// TwinCAT 3 PLC project Biegbert_SPS
// ProgramVersion: 3.1.4026.27
// CompilerDefines: SIM
// libraries:
//   Tc2_MC2, * (Beckhoff Automation GmbH)
//   Tc2_MC2_Camming, * (Beckhoff Automation GmbH)
//   Tc2_Standard, * (Beckhoff Automation GmbH)
//   Tc2_System, * (Beckhoff Automation GmbH)
//   TcUnit, * (www.tcunit.org)
// project tree:
//   07_Test/ FB_BendKinematics_Test.TcPOU, PRG_TEST.TcPOU
//   00_GVL/ GVL_Config.TcGVL, GVL_HMI.TcGVL, GVL_Axis.TcGVL, GVL_Devices.TcGVL, GVL_IO.TcGVL, GVL_Plan.TcGVL, GVL_Sim.TcGVL
//   01_DUT/ E_AlarmCode.TcDUT, E_AlarmSeverity.TcDUT, E_Axis.TcDUT, E_AxisState.TcDUT, E_ClampState.TcDUT, E_CmdResult.TcDUT, E_HmiCmd.TcDUT, E_KinState.TcDUT, E_MotionMode.TcDUT, E_OperatingMode.TcDUT, ST_AlarmEntry.TcDUT, ST_HmiAlarms.TcDUT, ST_HmiAxisStatus.TcDUT, ST_HmiClampStatus.TcDUT, ST_HmiCmd.TcDUT, ST_HmiCmdAck.TcDUT, ST_HmiIoStatus.TcDUT, ST_HmiJog.TcDUT, ST_HmiParam.TcDUT, ST_HmiStatus.TcDUT, ST_KinStatus.TcDUT, ST_Material.TcDUT, E_G0Step.TcDUT, E_G2Step.TcDUT, E_G3Step.TcDUT, ST_FeedPoint.TcDUT, ST_PlanHeader.TcDUT, ST_PlanPoint.TcDUT, ST_PlanSection.TcDUT, ST_PlanTransfer.TcDUT, ST_RotPoint.TcDUT
//   04_Kinematics/ FB_BendKinematics.TcPOU, I_Kinematics.TcIO, F_ChuckInZone.TcPOU, F_ClampBlocking.TcPOU, F_Z1Max.TcPOU
//   02_IO/ FB_IoMap.TcPOU, FB_IoSim.TcPOU
//   03_Devices/ FB_Axis.TcPOU, FB_Clamp.TcPOU, F_Mod360.TcPOU
//   05_Sequence/ FB_BendSequence.TcPOU, FB_Interlocks.TcPOU, FB_ModeManager.TcPOU
//   06_HMI/ FB_AlarmManager.TcPOU, FB_HmiCommand.TcPOU, FB_HmiStatus.TcPOU, FB_PlanStore.TcPOU, F_PlanChecksum.TcPOU
//   / PlcTask.TcTTO
//   POUs/ MAIN.TcPOU
// real-time tasks:
//   TASK PlcTask: cycle T#10ms, priority 20, ADS port 350
// motion (NC):
//   TASK NC-Task 1 SAF: cycle T#2ms, priority 4, ADS port 501
//   TASK NC-Task 1 SVB: cycle T#10ms, priority 8, ADS port 511
//   AXIS Z1 (id 1)
//     Dynamic: AccelerationMaximum=200, DecelerationMaximum=200, Acceleration=200, Deceleration=200
//     Velo: Maximum=50
//     OtherSettings: AllowMotionCmdToSlave=true
//     encoder EncType=1
//       SoftEndMinControl: Enable=true, Range=-30
//       SoftEndMaxControl: Enable=true, Range=1282
//     drive DrvType=5
//       Analog: VeloReferenz=100, TorqueSetpointScale=10, ScaleFactorActTorque=0.1
//       TimeComp: TaskDelayCycles=1
//     controller CtrType=1
//       CtrPara: PriorControlFactor=1
//         Observer: BandWidth=20
//   AXIS Z2 (id 2)
//     Dynamic: AccelerationMaximum=100, DecelerationMaximum=100, Acceleration=100, Deceleration=100
//     Velo: Maximum=28.6
//     OtherSettings: AllowMotionCmdToSlave=true
//     encoder EncType=1
//       SoftEndMinControl: Enable=true, Range=-50
//       SoftEndMaxControl: Enable=true, Range=48
//     drive DrvType=5
//       Analog: VeloReferenz=57.2, TorqueSetpointScale=10, ScaleFactorActTorque=0.1
//     controller CtrType=1
//       CtrPara: PriorControlFactor=1
//         Observer: BandWidth=20
//   AXIS X (id 3)
//     Dynamic: AccelerationMaximum=20, DecelerationMaximum=20, Acceleration=20, Deceleration=20
//     Velo: Maximum=3.5
//     OtherSettings: AllowMotionCmdToSlave=true
//     encoder EncType=1
//       SoftEndMinControl: Enable=true, Range=-50
//       SoftEndMaxControl: Enable=true, Range=50
//     drive DrvType=5
//       Analog: VeloReferenz=7, TorqueSetpointScale=10, ScaleFactorActTorque=0.1
//     controller CtrType=1
//       CtrPara: PriorControlFactor=1
//         Observer: BandWidth=20
//   AXIS A (id 4)
//     General: UnitName=°
//     Dynamic: AccelerationMaximum=360, DecelerationMaximum=360, Acceleration=360, Deceleration=360
//     Velo: Maximum=180
//     OtherSettings: AllowMotionCmdToSlave=true
//     encoder EncType=1
//       SoftEndMinControl: Enable=true, Range=-60
//       SoftEndMaxControl: Enable=true, Range=60
//     drive DrvType=5
//       Analog: VeloReferenz=360, TorqueSetpointScale=10, ScaleFactorActTorque=0.1
//     controller CtrType=1
//       CtrPara: PriorControlFactor=1
//         Observer: BandWidth=20
//   AXIS W (id 5)
//     Dynamic: AccelerationMaximum=360, DecelerationMaximum=360, Acceleration=360, Deceleration=360
//     Velo: Maximum=180
//     OtherSettings: AllowMotionCmdToSlave=true
//     encoder EncType=1
//     drive DrvType=5
//       Analog: VeloReferenz=360, TorqueSetpointScale=10, ScaleFactorActTorque=0.1
//     controller CtrType=1
//       CtrPara: PriorControlFactor=1
//         Observer: BandWidth=20
// variable links:
//   (this object) <-> NC-Task 1 SAF/Axes/A
//     PlcTask Inputs/GVL_Axis.A.NcToPlc <-> Outputs/ToPlc
//     PlcTask Outputs/GVL_Axis.A.PlcToNc <-> Inputs/FromPlc
//   (this object) <-> NC-Task 1 SAF/Axes/W
//     PlcTask Inputs/GVL_Axis.W.NcToPlc <-> Outputs/ToPlc
//     PlcTask Outputs/GVL_Axis.W.PlcToNc <-> Inputs/FromPlc
//   (this object) <-> NC-Task 1 SAF/Axes/X
//     PlcTask Inputs/GVL_Axis.X.NcToPlc <-> Outputs/ToPlc
//     PlcTask Outputs/GVL_Axis.X.PlcToNc <-> Inputs/FromPlc
//   (this object) <-> NC-Task 1 SAF/Axes/Z1
//     PlcTask Inputs/GVL_Axis.Z1.NcToPlc <-> Outputs/ToPlc
//     PlcTask Outputs/GVL_Axis.Z1.PlcToNc <-> Inputs/FromPlc
//   (this object) <-> NC-Task 1 SAF/Axes/Z2
//     PlcTask Inputs/GVL_Axis.Z2.NcToPlc <-> Outputs/ToPlc
//     PlcTask Outputs/GVL_Axis.Z2.PlcToNc <-> Inputs/FromPlc

CONFIGURATION Biegbert_SPS
    RESOURCE PLC ON TwinCAT3
        TASK PlcTask(INTERVAL := T#10ms, PRIORITY := 20);
        PROGRAM MAIN WITH PlcTask : MAIN;
    END_RESOURCE
END_CONFIGURATION

// ---- 01_DUT/E_AlarmCode.TcDUT
// Alarmcodes. Die Texte liegen im Backend (backend/biegbert/alarms.py).
{attribute 'qualified_only'}
{attribute 'strict'}
{attribute 'to_string'}
TYPE E_AlarmCode :
(
    None := 0,
    HmiHeartbeatLost := 1001, // Heartbeat ausgefallen
    SimulationActive := 1002, // Simulationsbetrieb aktiv
    EStopActive := 1100, // Not-Halt ausgelöst
    SafetyNotReady := 1101, // TwinSAFE nicht betriebsbereit
    AxisError := 2000, // nSource = E_Axis, nDetail = NC-Fehlercode
    AxisLagError := 2001, // Schleppfehler
    AxisSoftLimit := 2002, // Software-Endlage
    AxisTorqueLimit := 2003, // Momentgrenze
    ClampTimeout := 3000, // nSource = Niederhalter
    ClampPressureLow := 3001, // Klemmdruck fehlt
    ClampZoneViolation := 3002, // 4BF-Zone bei geschlossenem Niederhalter
    DistanceZ1Z2 := 4000, // dZ12 unterschritten
    KinCoupleFailed := 5000, // Kopplung oder Kurvenscheibe fehlgeschlagen, nDetail = NC-Fehlercode
    KinMasterFault := 5001, // Master Z1 gestört
    KinSlaveFault := 5002, // Slave gestört
    KinPositionDeviation := 5003, // Achse weicht vor Wiederanlauf vom Plan ab
    SeqStepTimeout := 6001 // Schritt hängt, nDetail = Schrittnummer
) UDINT;
END_TYPE

// ---- 01_DUT/E_AlarmSeverity.TcDUT
// Abgestufte Reaktion nach SE3.
{attribute 'qualified_only'}
{attribute 'strict'}
{attribute 'to_string'}
TYPE E_AlarmSeverity :
(
    None := 0,
    Info := 1, // nur Anzeige
    Warning := 2, // Anzeige, Ablauf läuft weiter
    Stop := 3, // Pause
    Fault := 4 // Pause, Wiederanlauf erst nach Behebung
) INT;
END_TYPE

// ---- 01_DUT/E_Axis.TcDUT
// Achsen. Die Werte sind die Indizes von aAxis in ST_HmiStatus.
{attribute 'qualified_only'}
{attribute 'strict'}
{attribute 'to_string'}
TYPE E_Axis :
(
    None := 0, // keine Achse
    Z1 := 1, // Vorschub, mm
    Z2 := 2, // Führung, mm
    X := 3, // Matrizenauslenkung, mm
    A := 4, // Matrizendrehung, °
    W := 5 // Rohrdrehung, °, Modulo
) INT;
END_TYPE

// ---- 01_DUT/E_AxisState.TcDUT
// Vereinfachter Achszustand für die GUI.
{attribute 'qualified_only'}
{attribute 'strict'}
{attribute 'to_string'}
TYPE E_AxisState :
(
    Disabled := 0,
    Standstill := 1,
    Moving := 2, // Einzelbewegung
    Coupled := 3, // über FB_BendKinematics gekoppelt
    Error := 4
) INT;
END_TYPE

// ---- 01_DUT/E_ClampState.TcDUT
// Zustand eines Niederhalters.
{attribute 'qualified_only'}
{attribute 'strict'}
{attribute 'to_string'}
TYPE E_ClampState :
(
    Unknown := 0,
    Open := 1, // Endlage OFFEN gemeldet
    Closing := 2, // Ventil an, Schaltzeit läuft
    Clamped := 3, // OFFEN verlassen, Druck ok, Schaltzeit abgelaufen
    Opening := 4, // Ventil aus, Endlage noch nicht erreicht
    Fault := 5 // Zeitüberwachung oder Plausibilität verletzt
) INT;
END_TYPE

// ---- 01_DUT/E_CmdResult.TcDUT
// Ergebnis der Kommandoprüfung.
{attribute 'qualified_only'}
{attribute 'strict'}
{attribute 'to_string'}
TYPE E_CmdResult :
(
    None := 0, // noch keine Antwort
    Accepted := 1, // angenommen, Ausführung siehe Status
    RejectedUnknown := 2, // Kommando unbekannt
    RejectedMode := 3, // in dieser Betriebsart nicht erlaubt
    RejectedInterlock := 4, // Verriegelung aktiv
    RejectedParam := 5, // Parameter ungültig
    RejectedSequence := 6, // zweite Stufe ohne gültige erste Stufe
    RejectedBusy := 7 // Gerät beschäftigt
) INT;
END_TYPE

// ---- 01_DUT/E_HmiCmd.TcDUT
// Kommandos der GUI. Details: docs/hmi-schnittstelle.md
{attribute 'qualified_only'}
{attribute 'strict'}
{attribute 'to_string'}
TYPE E_HmiCmd :
(
    None := 0,
    AlarmAck := 10, // nValue = Alarm-Slot, 0 = alle
    ParamApply := 11, // stParam prüfen und übernehmen
    AxisEnable := 100, // Phase 4/6: eAxis
    AxisDisable := 101, // Phase 6: eAxis
    AxisReset := 102, // Phase 6: eAxis
    AxisHalt := 103, // Phase 4/6: eAxis
    AxisMoveAbs := 104, // Phase 6: eAxis, fPosition, fVelocity
    ClampOpen := 120, // Phase 6: nClamp
    ClampClose := 121, // Phase 6: nClamp
    ModePause := 200, // Phase 6
    ModeResume1 := 201, // Phase 6: RES1
    ModeResume2 := 202, // Phase 6: RES2
    ModeSingleAxis1 := 203, // Phase 6: MAN1
    ModeSingleAxis2 := 204, // Phase 6: MAN2
    ModeReturnToBase := 205, // Phase 6: OK, nur bei GZ_POS
    SimSetInput := 300, // Phase 5/6: nur im Simulationsbetrieb, nValue = Signal-ID, fPosition <> 0 = TRUE
    SimInjectFault := 301, // Phase 5: nur im Simulationsbetrieb, nValue = Fehler-ID
    SeqStart := 400, // reserviert Phase 8: ST
    SeqConfirmQ1 := 401, // reserviert Phase 8
    SeqConfirmQ2 := 402, // reserviert Phase 8
    SeqPartRemoved := 403, // reserviert Phase 8: ENT
    PlanLoad := 410, // reserviert Phase 9
    MaterialConfirm := 411, // reserviert Phase 9
    CalibrateAxis := 500 // reserviert Phase 9: Einmessen
) UDINT;
END_TYPE

// ---- 01_DUT/E_KinState.TcDUT
// Zustand der Kinematik.
{attribute 'qualified_only'}
{attribute 'strict'}
{attribute 'to_string'}
TYPE E_KinState :
(
    Idle := 0, // kein Plan aktiv
    Loaded := 1, // Plan geladen, entkoppelt
    Coupling := 2,
    Running := 3, // gekoppelt, Master läuft
    Holding := 4, // Master bremst
    Held := 5, // gekoppelt, Stillstand
    Decoupling := 6,
    Fault := 7 // Reset nötig
) INT;
END_TYPE

// ---- 01_DUT/E_MotionMode.TcDUT
// Bewegungsmodus der Kinematik.
{attribute 'qualified_only'}
{attribute 'strict'}
{attribute 'to_string'}
TYPE E_MotionMode :
(
    Single := 1, // entkoppelt, Einzelachsen erlaubt
    Coupled := 2, // gekoppelt, Master läuft oder fährt an
    Hold := 3 // gekoppelt, Master hält
) INT;
END_TYPE

// ---- 01_DUT/E_OperatingMode.TcDUT
// Betriebsart. Die Werte entsprechen den GRAFCET-Schritten von G1.
{attribute 'qualified_only'}
{attribute 'strict'}
{attribute 'to_string'}
TYPE E_OperatingMode :
(
    Automatic := 10, // G1 Schritt 10
    Pause := 11, // G1 Schritt 11
    SingleAxis := 12, // G1 Schritt 12
    ReturnToBase := 13 // G1 Schritt 13
) INT;
END_TYPE

// ---- 01_DUT/ST_AlarmEntry.TcDUT
// Ein Alarm. Texte und Historie liegen im Backend.
{attribute 'pack_mode' := '1'}
TYPE ST_AlarmEntry :
STRUCT
    eCode : E_AlarmCode;
    eSeverity : E_AlarmSeverity;
    nSource : DINT; // Achse oder Niederhalter
    nDetail : UDINT;
    nTimestamp : ULINT; // Windows-Dateizeit, 100 ns
    bActive : BOOL; // Ursache besteht noch
    bAcked : BOOL;
END_STRUCT
END_TYPE

// ---- 01_DUT/ST_HmiAlarms.TcDUT
// SPS -> GUI. Aktive oder nicht quittierte Alarme.
{attribute 'pack_mode' := '1'}
TYPE ST_HmiAlarms :
STRUCT
    nChangeCounter : UDINT; // bei jeder Änderung +1
    nCount : UINT;
    bOverflow : BOOL;
    eHighestSeverity : E_AlarmSeverity;
    aEntry : ARRAY[1..32] OF ST_AlarmEntry;
END_STRUCT
END_TYPE

// ---- 01_DUT/ST_HmiAxisStatus.TcDUT
// SPS -> GUI. Status einer Achse.
{attribute 'pack_mode' := '1'}
TYPE ST_HmiAxisStatus :
STRUCT
    eState : E_AxisState;
    bEnabled : BOOL;
    bReady : BOOL;
    bError : BOOL;
    nErrorId : UDINT;
    fActPos : LREAL; // mm oder °
    fSetPos : LREAL;
    fActVelo : LREAL; // mm/s oder °/s
    fSetVelo : LREAL;
    fLagError : LREAL; // mm oder °
    fTorque_Nm : LREAL;
END_STRUCT
END_TYPE

// ---- 01_DUT/ST_HmiClampStatus.TcDUT
// SPS -> GUI. Status eines Niederhalters.
{attribute 'pack_mode' := '1'}
TYPE ST_HmiClampStatus :
STRUCT
    eState : E_ClampState;
    bValve : BOOL; // Ausgang
    bOpen : BOOL; // Endlage OFFEN
    fLastSwitchTime_ms : LREAL;
END_STRUCT
END_TYPE

// ---- 01_DUT/ST_HmiCmd.TcDUT
// GUI -> SPS. Die GUI schreibt hier, die SPS liest nur.
{attribute 'pack_mode' := '1'}
TYPE ST_HmiCmd :
STRUCT
    nHeartbeat : UDINT; // alle 100 ms hochzählen
    nCmdId : UDINT; // zuletzt und getrennt schreiben
    eCmd : E_HmiCmd;
    eAxis : E_Axis;
    nClamp : USINT; // 1..6, 0 = keiner
    fPosition : LREAL; // mm oder °, je nach Achse
    fVelocity : LREAL; // mm/s oder °/s
    nValue : DINT; // kommandoabhängig
    stJog : ST_HmiJog;
END_STRUCT
END_TYPE

// ---- 01_DUT/ST_HmiCmdAck.TcDUT
// SPS -> GUI. Antwort auf das letzte Kommando.
{attribute 'pack_mode' := '1'}
TYPE ST_HmiCmdAck :
STRUCT
    nAckId : UDINT; // gleich nCmdId, sobald geprüft
    eResult : E_CmdResult;
    nDetail : UDINT; // z. B. fehlende Bedingung
END_STRUCT
END_TYPE

// ---- 01_DUT/ST_HmiIoStatus.TcDUT
// SPS -> GUI. E/A-Übersicht ohne Niederhalter. Belegung folgt mit der EMSR-Liste.
{attribute 'pack_mode' := '1'}
TYPE ST_HmiIoStatus :
STRUCT
    bPressureOk : BOOL; // Druckschalter SDE5
    abPanelIn : ARRAY[1..16] OF BOOL; // ED1809
    abPanelOut : ARRAY[1..16] OF BOOL; // ED2809
END_STRUCT
END_TYPE

// ---- 01_DUT/ST_HmiJog.TcDUT
// Tippen. Wird zyklisch ausgewertet und läuft nicht über den Handshake.
{attribute 'pack_mode' := '1'}
TYPE ST_HmiJog :
STRUCT
    eAxis : E_Axis;
    nDirection : SINT; // -1, 0, +1
    fVelocityFactor_pct : LREAL; // 0..100 der Einrichtgeschwindigkeit
END_STRUCT
END_TYPE

// ---- 01_DUT/ST_HmiParam.TcDUT
// GUI -> SPS mit Übernahme durch ParamApply.
{attribute 'pack_mode' := '1'}
TYPE ST_HmiParam :
STRUCT
    nPlanId : UDINT;
    stMaterial : ST_Material;
    fFeedOverride_pct : LREAL; // 0..100
    fSingleAxisVelo_pct : LREAL; // 0..100
END_STRUCT
END_TYPE

// ---- 01_DUT/ST_HmiStatus.TcDUT
// SPS -> GUI. Die SPS schreibt hier, die GUI liest nur.
{attribute 'pack_mode' := '1'}
TYPE ST_HmiStatus :
STRUCT
    nLifeCounter : UDINT; // pro SPS-Zyklus +1
    bHmiAlive : BOOL;
    bSimulation : BOOL;
    bEStopActive : BOOL;
    bSafetyOk : BOOL;
    eMode : E_OperatingMode;
    nStepG2 : INT; // GRAFCET-Schritt
    nStepG3 : INT;
    nBend : UDINT; // aktueller Bogen
    dwBaseStateMissing : DWORD; // Bitmaske, siehe Doku
    stCmdAck : ST_HmiCmdAck;
    aAxis : ARRAY[1..5] OF ST_HmiAxisStatus; // Index = E_Axis
    aClamp : ARRAY[1..6] OF ST_HmiClampStatus;
    stIo : ST_HmiIoStatus;
    stKin : ST_KinStatus;
    stParamActive : ST_HmiParam;
END_STRUCT
END_TYPE

// ---- 01_DUT/ST_KinStatus.TcDUT
// Status von I_Kinematics.
{attribute 'pack_mode' := '1'}
TYPE ST_KinStatus :
STRUCT
    eState : E_KinState;
    eMode : E_MotionMode;
    nPlanId : UDINT;
    bError : BOOL;
    nErrorId : UDINT;
    fMasterPos_mm : LREAL;
END_STRUCT
END_TYPE

// ---- 01_DUT/ST_Material.TcDUT
// Halbzeugdaten des aktiven Programms.
{attribute 'pack_mode' := '1'}
TYPE ST_Material :
STRUCT
    fDiameter_mm : LREAL;
    fWall_mm : LREAL; // 0 = Vollmaterial
    fYield_MPa : LREAL; // Rp0,2
    fForceLimit_N : LREAL;
END_STRUCT
END_TYPE

// ---- 01_DUT/E_G0Step.TcDUT
// GRAFCET G0 Not-Halt [Langfeld].
{attribute 'qualified_only'}
{attribute 'strict'}
{attribute 'to_string'}
TYPE E_G0Step :
(
    S1_Betrieb := 1,
    S2_NotHalt := 2
) INT;
END_TYPE

// ---- 01_DUT/E_G2Step.TcDUT
// GRAFCET G2 Biegevorgang [Langfeld], Nummern = GRAFCET-Schritte.
{attribute 'qualified_only'}
{attribute 'strict'}
{attribute 'to_string'}
TYPE E_G2Step :
(
    S20_Grundzustand := 20,      // wartet auf Start
    S21_Startposition := 21,     // Z2, X, A und Z1 auf Startposition des Abschnitts
    S22_Niederhalter := 22,      // NH_soll schließen, Klemmung prüfen
    S23_Biegen := 23,            // gekoppelt: Z1 Master, X und A aus Kurvenscheibe
    S24_Halten := 24,            // Geometrie unter Last halten, warten auf Q1
    S25_NhOeffnen := 25,         // alle Niederhalter öffnen, warten auf Q2
    S26_Neutral := 26,           // entkoppeln, X und A auf 0
    S27_Uebergabe := 27,         // n := n + 1; weiterer Abschnitt oder warten auf ENT / Fortsetzung
    S28_Grundstellung := 28      // Z1, Z2, W auf 0
) INT;
END_TYPE

// ---- 01_DUT/E_G3Step.TcDUT
// GRAFCET G3 Werkstückrotation [Langfeld].
{attribute 'qualified_only'}
{attribute 'strict'}
{attribute 'to_string'}
TYPE E_G3Step :
(
    S30_Bereit := 30,
    S31_Stop := 31,     // Master steht an der Rotationsposition
    S32_Drehen := 32    // W dreht
) INT;
END_TYPE

// ---- 01_DUT/ST_FeedPoint.TcDUT
// Ab Z1-Position fZ1_mm gilt der Vorschub fFeed_mm_s.
{attribute 'pack_mode' := '1'}
TYPE ST_FeedPoint :
STRUCT
    fZ1_mm : LREAL;
    fFeed_mm_s : LREAL;
END_STRUCT
END_TYPE

// ---- 01_DUT/ST_PlanHeader.TcDUT
{attribute 'pack_mode' := '1'}
TYPE ST_PlanHeader :
STRUCT
    nPlanId : UDINT;
    nFormat : UINT;           // = GVL_Config.cPlanFormat
    nSectionCount : UINT;
    nPointCount : UDINT;
    nChecksum : UDINT;        // F_PlanChecksum über die belegten Abschnitte und Punkte
    stMaterial : ST_Material;
END_STRUCT
END_TYPE

// ---- 01_DUT/ST_PlanPoint.TcDUT
// Stützpunkt der Kurvenscheibe: Masterposition s (= Z1) mit u (= X) und phi (= A).
{attribute 'pack_mode' := '1'}
TYPE ST_PlanPoint :
STRUCT
    fS_mm : LREAL;
    fU_mm : LREAL;
    fPhi_deg : LREAL;
END_STRUCT
END_TYPE

// ---- 01_DUT/ST_PlanSection.TcDUT
// Ein Abschnitt = eine Kurvenscheibe mit konstantem Z2. Geraden sind Teil der Kurvenscheibe (u = 0).
{attribute 'pack_mode' := '1'}
TYPE ST_PlanSection :
STRUCT
    fZ1Start_mm : LREAL;
    fZ1Fin_mm : LREAL;
    fZ2_mm : LREAL;
    nFirstPoint : UDINT;      // Index in aPoint (1-basiert)
    nPointCount : UDINT;
    nFeedCount : UINT;
    aFeed : ARRAY[1..8] OF ST_FeedPoint;     // = GVL_Config.cMaxFeed
    nRotCount : UINT;
    aRot : ARRAY[1..16] OF ST_RotPoint;      // = GVL_Config.cMaxRot
    nClampMask : BYTE;        // Bit 0..5: NH1..NH6 zu Beginn schließen
    aClampOpen_mm : ARRAY[1..6] OF LREAL;    // Z1-Position, ab der NH i geöffnet wird
END_STRUCT
END_TYPE

// ---- 01_DUT/ST_PlanTransfer.TcDUT
// Übergabebereich Biegeplan (GVL_HMI.stPlanXfer) und aktiver Plan (GVL_Plan.stActive). 103552 Byte.
{attribute 'pack_mode' := '1'}
TYPE ST_PlanTransfer :
STRUCT
    stHeader : ST_PlanHeader;
    aSection : ARRAY[1..16] OF ST_PlanSection;    // = GVL_Config.cMaxSections
    aPoint : ARRAY[1..4000] OF ST_PlanPoint;      // = GVL_Config.cMaxPoints
END_STRUCT
END_TYPE

// ---- 01_DUT/ST_RotPoint.TcDUT
// Rotation von W um fW_deg (relativ), wenn Z1 fZ1_mm erreicht.
{attribute 'pack_mode' := '1'}
TYPE ST_RotPoint :
STRUCT
    fZ1_mm : LREAL;
    fW_deg : LREAL;
END_STRUCT
END_TYPE

// ---- 00_GVL/GVL_Config.TcGVL
// Feste Konfigurationswerte. Werte mit VORLÄUFIG stammen aus Doku/CAD und werden an der Anlage ersetzt.
// Gleiche Werte stehen im Backend in backend/biegbert/config.py (siehe 04_Datenfluss_und_Zustaende, Kap. 6).
{attribute 'qualified_only'}
VAR_GLOBAL CONSTANT
    cAxisCount           : INT  := 5;
    cClampCount          : INT  := 6;
    cAlarmSlots          : INT  := 32;
    tHeartbeatTimeout    : TIME := T#500MS;
    tTwoStepConfirmation : TIME := T#10S;

    // Achsen, Index = E_Axis (1 Z1, 2 Z2, 3 X, 4 A, 5 W). VORLÄUFIG.
    // W ist in der NC eine Rundachse OHNE Modulo; die SPS rechnet die Anzeige auf 0..360°.
    aAxisMin        : ARRAY[1..5] OF LREAL := [-30.0, -50.0, -50.0, -60.0, -1.0E9];
    aAxisMax        : ARRAY[1..5] OF LREAL := [1282.0, 48.0, 50.0, 60.0, 1.0E9];
    aAxisVMax       : ARRAY[1..5] OF LREAL := [50.0, 28.6, 3.5, 180.0, 180.0];   // mm/s bzw. °/s
    aAxisVSetup     : ARRAY[1..5] OF LREAL := [30.0, 10.0, 3.5, 20.0, 30.0];    // Einrichtgeschwindigkeit bei 100 %
    aAxisAccel      : ARRAY[1..5] OF LREAL := [200.0, 100.0, 20.0, 360.0, 360.0];
    aRatedTorque_Nm : ARRAY[1..5] OF LREAL := [15.2, 1.2, 1.37, 2.38, 1.37];  // Motor-Nennmoment (Bezug von 0x6077), VORLÄUFIG
    fPosTol         : LREAL := 0.05;   // mm bzw. °

    // Prozessgeometrie (CAD-Auswertung 24.11.2026). VORLÄUFIG.
    fVAtZ2Zero_mm       : LREAL := 24.0;     // Werkzeugabstand v bei Z2 = 0
    fZ1CollisionBase_mm : LREAL := 743.25;   // Z1-Grenze Futter <-> Führung bei Z2 = 0
    // Z1-Bereich, in dem das Futter die Zone des Niederhalterpaares 1..3 berührt (Paar k = NH 2k-1, 2k)
    aClampZoneLo_mm : ARRAY[1..3] OF LREAL := [508.25, 278.5, 50.5];
    aClampZoneHi_mm : ARRAY[1..3] OF LREAL := [710.75, 481.0, 253.0];
    tClampSwitchSim : TIME := T#120MS;   // Schaltzeit im Simulationsmodell
    tClampSwitch    : TIME := T#120MS;   // Mindestzeit bis „geklemmt“ (DFM-50, an der Anlage messen)
    tClampTimeout   : TIME := T#1S;      // Zeitüberwachung Öffnen/Schließen

    fForceLimitMax_N : LREAL := 25000.0;

    // Planübergabe (muss zu backend/biegbert/plc/layout.py passen)
    cPlanFormat  : UINT := 1;
    cMaxSections : INT := 16;
    cMaxFeed     : INT := 8;
    cMaxRot      : INT := 16;
    cMaxPoints   : INT := 4000;
END_VAR

// ---- 00_GVL/GVL_HMI.TcGVL
// Einzige Schnittstelle zur GUI. Details: docs/hmi-schnittstelle.md
// Backend schreibt stCmd, stParam, stPlanXfer; die SPS schreibt stStatus und stAlarm.
{attribute 'qualified_only'}
VAR_GLOBAL
    stCmd      : ST_HmiCmd;
    stStatus   : ST_HmiStatus;
    stParam    : ST_HmiParam;
    stAlarm    : ST_HmiAlarms;
    stPlanXfer : ST_PlanTransfer;   // Übergabebereich Biegeplan, wird nur bei PlanLoad gelesen
END_VAR

// ---- 00_GVL/GVL_Axis.TcGVL
// NC-Achsen. Im System Manager unter MOTION > NC-Task > Achsen > (Achse) > Einstellungen > „Mit SPS verknüpfen“
// die passende Variable wählen: Z1 -> GVL_Axis.Z1 usw.
{attribute 'qualified_only'}
VAR_GLOBAL
    Z1 : AXIS_REF;   // Vorschub
    Z2 : AXIS_REF;   // Führung („Eisenschwein“)
    X  : AXIS_REF;   // Matrizenauslenkung
    A  : AXIS_REF;   // Matrizendrehung
    W  : AXIS_REF;   // Rohrdrehung
END_VAR

// ---- 00_GVL/GVL_Devices.TcGVL
// Geräteinstanzen. MAIN ruft sie zyklisch auf; Ablauf und HMI-Bausteine rufen nur ihre Methoden.
{attribute 'qualified_only'}
VAR_GLOBAL
    aAxis   : ARRAY[1..5] OF FB_Axis;    // Index = E_Axis
    aClamp  : ARRAY[1..6] OF FB_Clamp;
    fbKin   : FB_BendKinematics;
    fbAlarm : FB_AlarmManager;
END_VAR

// ---- 00_GVL/GVL_IO.TcGVL
// Prozessabbild und logische Signale. Nur 02_IO greift auf die AT-Variablen zu (architektur.md, Regel 5).
// Die AT-Variablen im System Manager mit den Klemmen verknüpfen (docs/twincat-einrichtung.md).
{attribute 'qualified_only'}
VAR_GLOBAL
    // ── Eingänge ──
    abClampOpenIn    AT %I* : ARRAY[1..6] OF BOOL;   // EP1008 Kanal 1..6: SMT-8M Endlage OFFEN, NH1..NH6
    bPressureOkIn    AT %I* : BOOL;                  // EP1008 Kanal 7: SDE5 Klemmdruck in Ordnung
    bSafetyOkIn      AT %I* : BOOL;                  // TwinSAFE -> Standard-SPS: Sicherheitskreis geschlossen, STO aufgehoben
    bEStopReleasedIn AT %I* : BOOL;                  // TwinSAFE -> Standard-SPS: Not-Halt entriegelt
    abPanelIn        AT %I* : ARRAY[1..16] OF BOOL;  // ED1809, Belegung offen
    anTorqueIn       AT %I* : ARRAY[1..5] OF INT;    // AX8000 Torque actual value (0x6077, 0,1 % Nennmoment), Index = E_Axis
    // ── Ausgänge ──
    abClampValveOut  AT %Q* : ARRAY[1..6] OF BOOL;   // EP2008 Kanal 1..6: Ventil NH1..NH6, TRUE = schließen
    abPanelOut       AT %Q* : ARRAY[1..16] OF BOOL;  // ED2809, Belegung offen
    bCameraTriggerOut AT %Q* : BOOL;                 // EL2252 Kanal 1 (später)

    // ── logische Signale (FB_IoMap) ──
    abClampOpen  : ARRAY[1..6] OF BOOL;
    bPressureOk  : BOOL;
    bSafetyOk    : BOOL;
    bEStopActive : BOOL;
    abPanel      : ARRAY[1..16] OF BOOL;
    afTorque_Nm  : ARRAY[1..5] OF LREAL;
    abClampValve : ARRAY[1..6] OF BOOL;
    abPanelLamp  : ARRAY[1..16] OF BOOL;
    bCameraTrigger : BOOL;
END_VAR

// ---- 00_GVL/GVL_Plan.TcGVL
// Geprüfte Kopie des aktiven Biegeplans. Schreibt nur FB_PlanStore, liest FB_BendKinematics und FB_BendSequence.
{attribute 'qualified_only'}
VAR_GLOBAL
    stActive : ST_PlanTransfer;
    bValid   : BOOL;
END_VAR

// ---- 00_GVL/GVL_Sim.TcGVL
// Eingriffe der Simulation. Wirkt nur, wenn das Projekt mit dem Compiler-Define SIM übersetzt wurde.
// Gesetzt über die Kommandos SimSetInput und SimInjectFault.
{attribute 'qualified_only'}
VAR_GLOBAL
    bPressureOk  : BOOL := TRUE;
    bEStop       : BOOL;
    abAxisFault  : ARRAY[1..5] OF BOOL;   // simulierter Achsfehler, Index = E_Axis
    abClampStuck : ARRAY[1..6] OF BOOL;   // Endlage OFFEN bleibt hängen
END_VAR

// ---- 04_Kinematics/I_Kinematics.TcIO
// Einzige Schnittstelle des Ablaufs zur Achskopplung. Details: docs/kinematik.md
INTERFACE I_Kinematics

METHOD Cyclic
// Einmal pro SPS-Zyklus aufrufen.
VAR_INPUT
END_VAR
END_METHOD

METHOD LoadPlan : BOOL
// Aktiven Plan (GVL_Plan.stActive) mit dieser ID übernehmen. Nur entkoppelt.
VAR_INPUT
    nPlanId : UDINT;
END_VAR
END_METHOD

METHOD LoadSection : BOOL
// Kurvenscheiben des Abschnitts nSection laden. Nur entkoppelt; fertig, wenn TableReady() TRUE meldet.
VAR_INPUT
    nSection : INT;
END_VAR
END_METHOD

METHOD TableReady : BOOL
VAR_INPUT
END_VAR
END_METHOD

METHOD Start : BOOL
// Koppelt X und A an Z1 und startet den Master.
VAR_INPUT
END_VAR
END_METHOD

METHOD Hold : BOOL
// Bremst den Master. Die Kopplung bleibt bestehen.
VAR_INPUT
END_VAR
END_METHOD

METHOD Resume : BOOL
// Setzt den Master aus dem Halt fort (nicht an einer offenen Rotation oder am Abschnittsende).
VAR_INPUT
END_VAR
END_METHOD

METHOD AtRotation : BOOL
// Master steht an einer Rotationsposition; RotationAngle() liefert den Drehwinkel für W.
VAR_INPUT
END_VAR
END_METHOD

METHOD RotationAngle : LREAL
VAR_INPUT
END_VAR
END_METHOD

METHOD ContinueAfterRotation : BOOL
VAR_INPUT
END_VAR
END_METHOD

METHOD SectionDone : BOOL
// Master steht am Ende des Abschnitts, Kopplung besteht noch.
VAR_INPUT
END_VAR
END_METHOD

METHOD Abort : BOOL
// Stoppt den Master und löst die Kopplung.
VAR_INPUT
END_VAR
END_METHOD

METHOD Reset : BOOL
// Quittiert einen Fehler der Kinematik. Der Plan bleibt erhalten.
VAR_INPUT
END_VAR
END_METHOD

METHOD Unload : BOOL
// Plan verwerfen (nur entkoppelt).
VAR_INPUT
END_VAR
END_METHOD

METHOD IsCoupled : BOOL
VAR_INPUT
END_VAR
END_METHOD

METHOD GetStatus : ST_KinStatus
VAR_INPUT
END_VAR
END_METHOD

END_INTERFACE

// ---- POUs/MAIN.TcPOU
PROGRAM MAIN
// Zyklusreihenfolge nach docs/architektur.md:
// 1 Eingänge, 2 Kommandos, 3 Abläufe, 4 Kinematik und Geräte, 5 Ausgänge, 6 Status und Alarme.
VAR
    fbIo : FB_IoMap;
    fbCmd : FB_HmiCommand;
    fbMode : FB_ModeManager;
    fbSeq : FB_BendSequence;
    fbPlan : FB_PlanStore;
    fbInterlocks : FB_Interlocks;
    fbStatus : FB_HmiStatus;
    dwBaseMissing : DWORD;
    bKinLock : BOOL;
    abSimFault : ARRAY[1..5] OF BOOL;
    bSim : BOOL;
    bInit : BOOL := TRUE;
    i : INT;
END_VAR

// 1 Eingänge
fbIo.ReadInputs();
bSim := fbIo.IsSimulation();
IF bInit THEN
    bInit := FALSE;
    IF bSim THEN
        GVL_Devices.fbAlarm.Raise(E_AlarmCode.SimulationActive, E_AlarmSeverity.Info, 0, 0);
    END_IF
END_IF
{IF defined (SIM)}
abSimFault := GVL_Sim.abAxisFault;
{END_IF}

// 2 Kommandos
dwBaseMissing := fbStatus.CalcBaseMissing(fbSeq.bMaterialOk);
fbCmd(fbMode := fbMode, fbSeq := fbSeq, fbPlan := fbPlan, dwBaseMissing := dwBaseMissing, bSimulation := bSim);

// 3 Abläufe
fbMode(bEStopActive := GVL_IO.bEStopActive, bSafetyOk := GVL_IO.bSafetyOk,
       nStopCounter := GVL_Devices.fbAlarm.nStopCounter);
fbSeq(bFree := fbMode.bFree, bAbort := fbMode.bEnteredSingle, bInit := fbMode.bInitSequences);

// 4 Kinematik und Geräte
GVL_Devices.fbKin.Cyclic();
bKinLock := GVL_Devices.fbKin.IsCoupled();
GVL_Devices.aAxis[1](pAxis := ADR(GVL_Axis.Z1), nIndex := 1, bAllowPower := NOT GVL_IO.bEStopActive,
    bLockedByKin := bKinLock, bSimFault := abSimFault[1], fTorque_Nm := GVL_IO.afTorque_Nm[1],
    fPowerOverride_pct := SEL(bKinLock, 100.0, GVL_HMI.stStatus.stParamActive.fFeedOverride_pct));
GVL_Devices.aAxis[2](pAxis := ADR(GVL_Axis.Z2), nIndex := 2, bAllowPower := NOT GVL_IO.bEStopActive,
    bLockedByKin := FALSE, bSimFault := abSimFault[2], fTorque_Nm := GVL_IO.afTorque_Nm[2]);
GVL_Devices.aAxis[3](pAxis := ADR(GVL_Axis.X), nIndex := 3, bAllowPower := NOT GVL_IO.bEStopActive,
    bLockedByKin := bKinLock, bSimFault := abSimFault[3], fTorque_Nm := GVL_IO.afTorque_Nm[3]);
GVL_Devices.aAxis[4](pAxis := ADR(GVL_Axis.A), nIndex := 4, bAllowPower := NOT GVL_IO.bEStopActive,
    bLockedByKin := bKinLock, bSimFault := abSimFault[4], fTorque_Nm := GVL_IO.afTorque_Nm[4]);
GVL_Devices.aAxis[5](pAxis := ADR(GVL_Axis.W), nIndex := 5, bAllowPower := NOT GVL_IO.bEStopActive,
    bLockedByKin := FALSE, bSimFault := abSimFault[5], fTorque_Nm := GVL_IO.afTorque_Nm[5]);
FOR i := 1 TO 6 DO
    GVL_Devices.aClamp[i](bSensorOpen := GVL_IO.abClampOpen[i], bPressureOk := GVL_IO.bPressureOk,
                          bForceOpen := GVL_IO.bEStopActive);
    GVL_IO.abClampValve[i] := GVL_Devices.aClamp[i].bValve;
END_FOR
fbInterlocks();

// 5 Ausgänge
fbIo.WriteOutputs();

// 6 Status und Alarme
fbStatus(fbMode := fbMode, fbSeq := fbSeq, bHmiAlive := fbCmd.bHmiAlive, bSimulation := bSim,
         dwBaseMissing := dwBaseMissing);
GVL_Devices.fbAlarm.WriteTo(GVL_HMI.stAlarm);

{IF defined (TEST)}
PRG_TEST();
{END_IF}

END_PROGRAM

// ---- 02_IO/FB_IoMap.TcPOU
// Einzige Stelle mit Zugriff auf das Prozessabbild (E4). Füllt die logischen Signale aus Hardware oder Simulation.
FUNCTION_BLOCK FB_IoMap
VAR
    fbSim : FB_IoSim;
    i : INT;
END_VAR

// Aufruf über ReadInputs() und WriteOutputs().

METHOD ReadInputs
VAR_INPUT
END_VAR
{IF defined (SIM)}
fbSim(abValve := GVL_IO.abClampValve);
GVL_IO.abClampOpen := fbSim.abClampOpen;
GVL_IO.bPressureOk := GVL_Sim.bPressureOk;
GVL_IO.bEStopActive := GVL_Sim.bEStop;
GVL_IO.bSafetyOk := NOT GVL_Sim.bEStop;
FOR i := 1 TO 16 DO
    GVL_IO.abPanel[i] := FALSE;
END_FOR
FOR i := 1 TO 5 DO
    GVL_IO.afTorque_Nm[i] := 0.0;
END_FOR
{ELSE}
GVL_IO.abClampOpen := GVL_IO.abClampOpenIn;
GVL_IO.bPressureOk := GVL_IO.bPressureOkIn;
GVL_IO.bEStopActive := NOT GVL_IO.bEStopReleasedIn;
GVL_IO.bSafetyOk := GVL_IO.bSafetyOkIn;
GVL_IO.abPanel := GVL_IO.abPanelIn;
FOR i := 1 TO 5 DO
    GVL_IO.afTorque_Nm[i] := INT_TO_LREAL(GVL_IO.anTorqueIn[i]) * 0.001 * GVL_Config.aRatedTorque_Nm[i];
END_FOR
{END_IF}
END_METHOD

METHOD WriteOutputs
VAR_INPUT
END_VAR
{IF defined (SIM)}
// keine Hardware: Ausgänge bleiben aus
FOR i := 1 TO 6 DO
    GVL_IO.abClampValveOut[i] := FALSE;
END_FOR
FOR i := 1 TO 16 DO
    GVL_IO.abPanelOut[i] := FALSE;
END_FOR
GVL_IO.bCameraTriggerOut := FALSE;
{ELSE}
GVL_IO.abClampValveOut := GVL_IO.abClampValve;
GVL_IO.abPanelOut := GVL_IO.abPanelLamp;
GVL_IO.bCameraTriggerOut := GVL_IO.bCameraTrigger;
{END_IF}
END_METHOD

METHOD IsSimulation : BOOL
VAR_INPUT
END_VAR
{IF defined (SIM)}
IsSimulation := TRUE;
{ELSE}
IsSimulation := FALSE;
{END_IF}
END_METHOD

END_FUNCTION_BLOCK

// ---- 02_IO/FB_IoSim.TcPOU
// Simulationsmodell der Peripherie (nur mit Compiler-Define SIM aktiv): Endlagen der Niederhalter folgen den Ventilen.
FUNCTION_BLOCK FB_IoSim
VAR_INPUT
    abValve : ARRAY[1..6] OF BOOL;
END_VAR
VAR_OUTPUT
    abClampOpen : ARRAY[1..6] OF BOOL;
END_VAR
VAR
    aTonLeave : ARRAY[1..6] OF TON;   // Endlage OFFEN wird kurz nach dem Schalten verlassen
    aTonOpen  : ARRAY[1..6] OF TON;   // Endlage OFFEN wird nach der Schaltzeit erreicht
    i : INT;
END_VAR

FOR i := 1 TO 6 DO
    aTonLeave[i](IN := abValve[i], PT := T#20MS);
    aTonOpen[i](IN := NOT abValve[i], PT := GVL_Config.tClampSwitchSim);
    IF GVL_Sim.abClampStuck[i] THEN
        abClampOpen[i] := TRUE;
    ELSIF aTonLeave[i].Q THEN
        abClampOpen[i] := FALSE;
    ELSIF aTonOpen[i].Q THEN
        abClampOpen[i] := TRUE;
    END_IF
END_FOR

END_FUNCTION_BLOCK

// ---- 06_HMI/FB_HmiCommand.TcPOU
// Heartbeat-Überwachung, Kommando-Handshake und Tippen (docs/hmi-schnittstelle.md).
// Jede neue nCmdId wird genau einmal geprüft; Antwort: eResult, nDetail und zuletzt nAckId.
// Accepted heißt nur „angenommen“; den Fortschritt zeigt stStatus.
FUNCTION_BLOCK FB_HmiCommand
VAR_IN_OUT
    fbMode : FB_ModeManager;
    fbSeq : FB_BendSequence;
    fbPlan : FB_PlanStore;
END_VAR
VAR_INPUT
    dwBaseMissing : DWORD;
    bSimulation : BOOL;
END_VAR
VAR_OUTPUT
    bHmiAlive : BOOL;
END_VAR
VAR
    bInit : BOOL := TRUE;
    nLastCmdId : UDINT;
    nLastHb : UDINT;
    bHbSeen : BOOL;
    tonHb : TON;
    eRes : E_CmdResult;
    nDetail : UDINT;
    nJogAxis : INT;
    i : INT;
END_VAR

IF bInit THEN
    bInit := FALSE;
    nLastCmdId := GVL_HMI.stCmd.nCmdId;
    nLastHb := GVL_HMI.stCmd.nHeartbeat;
    GVL_HMI.stStatus.stCmdAck.nAckId := nLastCmdId;
    GVL_HMI.stStatus.stParamActive.nPlanId := 0;
    GVL_HMI.stStatus.stParamActive.stMaterial.fDiameter_mm := 15.0;
    GVL_HMI.stStatus.stParamActive.stMaterial.fWall_mm := 2.0;
    GVL_HMI.stStatus.stParamActive.stMaterial.fYield_MPa := 300.0;
    GVL_HMI.stStatus.stParamActive.stMaterial.fForceLimit_N := 16000.0;
    GVL_HMI.stStatus.stParamActive.fFeedOverride_pct := 100.0;
    GVL_HMI.stStatus.stParamActive.fSingleAxisVelo_pct := 100.0;
END_IF

// ── Heartbeat: jede Änderung von nHeartbeat ist ein Lebenszeichen ──
IF GVL_HMI.stCmd.nHeartbeat <> nLastHb THEN
    nLastHb := GVL_HMI.stCmd.nHeartbeat;
    bHbSeen := TRUE;
    tonHb(IN := FALSE);
END_IF
tonHb(IN := TRUE, PT := GVL_Config.tHeartbeatTimeout);
IF bHmiAlive AND (tonHb.Q OR NOT bHbSeen) THEN
    bHmiAlive := FALSE;
    GVL_Devices.fbAlarm.Raise(E_AlarmCode.HmiHeartbeatLost, E_AlarmSeverity.Stop, 0, 0);
    FOR i := 1 TO 5 DO
        IF GVL_Devices.aAxis[i].bBusy AND NOT GVL_Devices.aAxis[i].bLockedByKin THEN
            GVL_Devices.aAxis[i].Halt();
        END_IF
    END_FOR
ELSIF NOT bHmiAlive AND bHbSeen AND NOT tonHb.Q THEN
    bHmiAlive := TRUE;
    GVL_Devices.fbAlarm.Clear(E_AlarmCode.HmiHeartbeatLost, 0, FALSE);
END_IF

// ── Kommando ──
IF GVL_HMI.stCmd.nCmdId <> nLastCmdId THEN
    nLastCmdId := GVL_HMI.stCmd.nCmdId;
    nDetail := 0;
    eRes := Execute();
    GVL_HMI.stStatus.stCmdAck.eResult := eRes;
    GVL_HMI.stStatus.stCmdAck.nDetail := nDetail;
    GVL_HMI.stStatus.stCmdAck.nAckId := nLastCmdId;   // zuletzt
END_IF

Jog();

METHOD PRIVATE Execute : E_CmdResult
VAR
    nAx : INT;
    fTarget, fVMax, fDelta : LREAL;
    nBlk : INT;
    stKin : ST_KinStatus;
    eMode : E_OperatingMode;
    dwNotReady : DWORD;
    bCoupled : BOOL;
END_VAR
nAx := TO_INT(GVL_HMI.stCmd.eAxis);
eMode := fbMode.eMode;
stKin := GVL_Devices.fbKin.GetStatus();
bCoupled := GVL_Devices.fbKin.IsCoupled();

CASE GVL_HMI.stCmd.eCmd OF
E_HmiCmd.AlarmAck:
    GVL_Devices.fbAlarm.Ack(GVL_HMI.stCmd.nValue);
    fbMode.Acknowledge();
    FOR i := 1 TO 6 DO
        IF NOT GVL_Devices.aClamp[i].IsCommandedClosed() THEN
            GVL_Devices.aClamp[i].ResetFault();
        END_IF
    END_FOR
    IF stKin.eState = E_KinState.Fault AND NOT GVL_Devices.fbAlarm.FaultActive() THEN
        IF GVL_Devices.fbKin.Reset() THEN
            fbSeq.AbortRun();
        END_IF
    END_IF
    Execute := E_CmdResult.Accepted;

E_HmiCmd.ParamApply:
    IF bCoupled THEN
        Execute := E_CmdResult.RejectedMode;
    ELSIF GVL_HMI.stParam.fFeedOverride_pct < 0.0 OR GVL_HMI.stParam.fFeedOverride_pct > 100.0
          OR GVL_HMI.stParam.fSingleAxisVelo_pct <= 0.0 OR GVL_HMI.stParam.fSingleAxisVelo_pct > 100.0
          OR GVL_HMI.stParam.stMaterial.fDiameter_mm <= 0.0 OR GVL_HMI.stParam.stMaterial.fForceLimit_N <= 0.0 THEN
        Execute := E_CmdResult.RejectedParam;
    ELSE
        GVL_HMI.stStatus.stParamActive := GVL_HMI.stParam;
        GVL_HMI.stStatus.stParamActive.stMaterial.fForceLimit_N :=
            MIN(GVL_HMI.stParam.stMaterial.fForceLimit_N, GVL_Config.fForceLimitMax_N);
        Execute := E_CmdResult.Accepted;
    END_IF

E_HmiCmd.AxisEnable, E_HmiCmd.AxisDisable, E_HmiCmd.AxisReset, E_HmiCmd.AxisHalt, E_HmiCmd.AxisMoveAbs:
    IF nAx < 1 OR nAx > 5 THEN
        Execute := E_CmdResult.RejectedParam;
        RETURN;
    END_IF
    CASE GVL_HMI.stCmd.eCmd OF
    E_HmiCmd.AxisEnable:      // Phase-4-Ausnahme: ohne Betriebsartenprüfung
        IF GVL_IO.bEStopActive OR NOT GVL_IO.bSafetyOk THEN
            Execute := E_CmdResult.RejectedInterlock;
            nDetail := 1100;
        ELSE
            GVL_Devices.aAxis[nAx].Enable();
            Execute := E_CmdResult.Accepted;
        END_IF
    E_HmiCmd.AxisDisable:
        IF GVL_Devices.aAxis[nAx].bLockedByKin THEN
            Execute := E_CmdResult.RejectedBusy;
        ELSE
            GVL_Devices.aAxis[nAx].Disable();
            Execute := E_CmdResult.Accepted;
        END_IF
    E_HmiCmd.AxisReset:
        IF eMode <> E_OperatingMode.SingleAxis AND eMode <> E_OperatingMode.Pause THEN
            Execute := E_CmdResult.RejectedMode;
        ELSE
            {IF defined (SIM)}
            GVL_Sim.abAxisFault[nAx] := FALSE;
            {END_IF}
            GVL_Devices.aAxis[nAx].Reset();
            GVL_Devices.fbAlarm.Clear(E_AlarmCode.AxisLagError, nAx, FALSE);
            Execute := E_CmdResult.Accepted;
        END_IF
    E_HmiCmd.AxisHalt:
        IF GVL_Devices.aAxis[nAx].bLockedByKin THEN
            GVL_Devices.fbKin.Hold();
        ELSE
            GVL_Devices.aAxis[nAx].Halt();
        END_IF
        Execute := E_CmdResult.Accepted;
    E_HmiCmd.AxisMoveAbs:
        IF eMode <> E_OperatingMode.SingleAxis THEN
            Execute := E_CmdResult.RejectedMode;
            RETURN;
        END_IF
        IF NOT GVL_Devices.aAxis[nAx].bReady THEN
            Execute := E_CmdResult.RejectedInterlock;
            nDetail := 1;
            RETURN;
        END_IF
        IF GVL_Devices.aAxis[nAx].bLockedByKin THEN
            Execute := E_CmdResult.RejectedBusy;
            RETURN;
        END_IF
        fVMax := GVL_Config.aAxisVSetup[nAx] * GVL_HMI.stStatus.stParamActive.fSingleAxisVelo_pct / 100.0;
        IF GVL_HMI.stCmd.fVelocity <= 0.0 OR GVL_HMI.stCmd.fVelocity > fVMax + 1.0E-9 THEN
            Execute := E_CmdResult.RejectedParam;
            nDetail := 2;
            RETURN;
        END_IF
        fTarget := GVL_HMI.stCmd.fPosition;
        IF nAx = 5 THEN     // W: kürzester Weg zur Anzeigeposition 0..360°
            fDelta := F_Mod360(fTarget - F_Mod360(GVL_Devices.aAxis[5].fActPos) + 180.0) - 180.0;
            fTarget := GVL_Devices.aAxis[5].fActPos + fDelta;
        ELSIF fTarget < GVL_Config.aAxisMin[nAx] OR fTarget > GVL_Config.aAxisMax[nAx] THEN
            Execute := E_CmdResult.RejectedParam;
            nDetail := 1;
            RETURN;
        END_IF
        IF nAx = 1 THEN
            IF fTarget > F_Z1Max(GVL_Devices.aAxis[2].fActPos) + 1.0E-9 THEN
                Execute := E_CmdResult.RejectedInterlock;
                nDetail := 4000;
                RETURN;
            END_IF
            nBlk := F_ClampBlocking(GVL_Devices.aAxis[1].fActPos, fTarget);
            IF nBlk <> 0 THEN
                Execute := E_CmdResult.RejectedInterlock;
                nDetail := 3002;
                RETURN;
            END_IF
        ELSIF nAx = 2 THEN
            IF GVL_Devices.aAxis[1].fActPos > F_Z1Max(fTarget) + 1.0E-9 THEN
                Execute := E_CmdResult.RejectedInterlock;
                nDetail := 4000;
                RETURN;
            END_IF
        END_IF
        GVL_Devices.aAxis[nAx].MoveAbs(fTarget, GVL_HMI.stCmd.fVelocity);
        Execute := E_CmdResult.Accepted;
    END_CASE

E_HmiCmd.ClampOpen, E_HmiCmd.ClampClose:
    IF eMode <> E_OperatingMode.SingleAxis THEN
        Execute := E_CmdResult.RejectedMode;
    ELSIF GVL_HMI.stCmd.nClamp < 1 OR GVL_HMI.stCmd.nClamp > 6 THEN
        Execute := E_CmdResult.RejectedParam;
    ELSIF GVL_HMI.stCmd.eCmd = E_HmiCmd.ClampClose THEN
        IF F_ChuckInZone((USINT_TO_INT(GVL_HMI.stCmd.nClamp) + 1) / 2, GVL_Devices.aAxis[1].fActPos) THEN
            Execute := E_CmdResult.RejectedInterlock;
            nDetail := 3002;
        ELSE
            GVL_Devices.aClamp[GVL_HMI.stCmd.nClamp].Close();
            Execute := E_CmdResult.Accepted;
        END_IF
    ELSE
        GVL_Devices.aClamp[GVL_HMI.stCmd.nClamp].Open();
        Execute := E_CmdResult.Accepted;
    END_IF

E_HmiCmd.ModePause:
    Execute := fbMode.CmdPause();
E_HmiCmd.ModeResume1, E_HmiCmd.ModeSingleAxis1:
    Execute := fbMode.CmdFirstStage(GVL_HMI.stCmd.eCmd);
E_HmiCmd.ModeResume2, E_HmiCmd.ModeSingleAxis2:
    Execute := fbMode.CmdSecondStage(GVL_HMI.stCmd.eCmd, bHmiAlive, FaultActive());
E_HmiCmd.ModeReturnToBase:
    Execute := fbMode.CmdReturnToBase(dwMissing := dwBaseMissing, nDetail => nDetail);

E_HmiCmd.SimSetInput, E_HmiCmd.SimInjectFault:
    {IF defined (SIM)}
    Execute := Simulate();
    {ELSE}
    Execute := E_CmdResult.RejectedMode;
    {END_IF}

E_HmiCmd.PlanLoad:
    IF NOT fbSeq.CanLoadPlan() OR bCoupled THEN
        Execute := E_CmdResult.RejectedBusy;
        RETURN;
    END_IF
    nDetail := fbPlan.Load(DINT_TO_UDINT(GVL_HMI.stCmd.nValue));
    IF nDetail <> 0 THEN
        Execute := E_CmdResult.RejectedParam;
        RETURN;
    END_IF
    IF NOT GVL_Devices.fbKin.LoadPlan(DINT_TO_UDINT(GVL_HMI.stCmd.nValue)) THEN
        Execute := E_CmdResult.RejectedBusy;
        RETURN;
    END_IF
    fbSeq.SetMaterial(FALSE);
    Execute := E_CmdResult.Accepted;

E_HmiCmd.MaterialConfirm:
    IF stKin.nPlanId = 0 OR stKin.nPlanId <> DINT_TO_UDINT(GVL_HMI.stCmd.nValue) THEN
        Execute := E_CmdResult.RejectedParam;
    ELSE
        fbSeq.SetMaterial(TRUE);
        Execute := E_CmdResult.Accepted;
    END_IF

E_HmiCmd.SeqStart:
    dwNotReady := 0;
    FOR i := 1 TO 5 DO
        IF NOT GVL_Devices.aAxis[i].bReady THEN
            dwNotReady := dwNotReady OR SHL(DWORD#1, i);
        END_IF
    END_FOR
    IF eMode <> E_OperatingMode.Automatic THEN
        Execute := E_CmdResult.RejectedMode;
    ELSIF stKin.eState <> E_KinState.Loaded OR NOT GVL_Plan.bValid THEN
        Execute := E_CmdResult.RejectedInterlock;
        nDetail := 16#100;
    ELSIF NOT fbSeq.bMaterialOk THEN
        Execute := E_CmdResult.RejectedInterlock;
        nDetail := 16#200;
    ELSIF GVL_IO.bEStopActive THEN
        Execute := E_CmdResult.RejectedInterlock;
        nDetail := 1100;
    ELSIF NOT bHmiAlive THEN
        Execute := E_CmdResult.RejectedInterlock;
        nDetail := 1001;
    ELSIF dwNotReady <> 0 THEN
        Execute := E_CmdResult.RejectedInterlock;
        nDetail := 16#10000 OR DWORD_TO_UDINT(dwNotReady);
    ELSIF FaultActive() THEN
        Execute := E_CmdResult.RejectedInterlock;
        nDetail := 16#40;
    ELSE
        Execute := fbSeq.Start(dwBaseMissing := dwBaseMissing, nDetail => nDetail);
    END_IF

E_HmiCmd.SeqConfirmQ1:
    Execute := fbSeq.ConfirmQ1();
E_HmiCmd.SeqConfirmQ2:
    Execute := fbSeq.ConfirmQ2();
E_HmiCmd.SeqPartRemoved:
    Execute := fbSeq.PartRemoved();

ELSE
    Execute := E_CmdResult.RejectedUnknown;   // CalibrateAxis und unbekannte Kommandos
END_CASE
END_METHOD

METHOD PRIVATE FaultActive : BOOL
VAR
    k : INT;
END_VAR
FaultActive := GVL_Devices.fbAlarm.FaultActive();
FOR k := 1 TO 5 DO
    IF GVL_Devices.aAxis[k].bError THEN
        FaultActive := TRUE;
    END_IF
END_FOR
END_METHOD

METHOD PRIVATE Simulate : E_CmdResult
// SimSetInput: nValue 1 Druckschalter, 2 Not-Halt; fPosition <> 0 = TRUE.
// SimInjectFault: 1 Achsfehler Z1, 2 X, 3 A, 4 Druckabfall, 5 Not-Halt, 6 Schleppfehler-Warnung Z1.
VAR
END_VAR
Simulate := E_CmdResult.Accepted;
IF GVL_HMI.stCmd.eCmd = E_HmiCmd.SimSetInput THEN
    CASE GVL_HMI.stCmd.nValue OF
    1: GVL_Sim.bPressureOk := GVL_HMI.stCmd.fPosition <> 0.0;
    2: GVL_Sim.bEStop := GVL_HMI.stCmd.fPosition <> 0.0;
    ELSE
        Simulate := E_CmdResult.RejectedParam;
    END_CASE
ELSE
    CASE GVL_HMI.stCmd.nValue OF
    1: GVL_Sim.abAxisFault[1] := TRUE;
    2: GVL_Sim.abAxisFault[3] := TRUE;
    3: GVL_Sim.abAxisFault[4] := TRUE;
    4: GVL_Sim.bPressureOk := FALSE;
    5: GVL_Sim.bEStop := TRUE;
    6: GVL_Devices.fbAlarm.Raise(E_AlarmCode.AxisLagError, E_AlarmSeverity.Warning, 1, 123);
    ELSE
        Simulate := E_CmdResult.RejectedParam;
    END_CASE
END_IF
END_METHOD

METHOD PRIVATE Jog
VAR
    nAx : INT;
    nDir : INT;
    bOk : BOOL;
    fVel : LREAL;
END_VAR
nAx := TO_INT(GVL_HMI.stCmd.stJog.eAxis);
nDir := SINT_TO_INT(GVL_HMI.stCmd.stJog.nDirection);
bOk := fbMode.eMode = E_OperatingMode.SingleAxis AND bHmiAlive AND (nDir = 1 OR nDir = -1) AND nAx >= 1 AND nAx <= 5;
IF bOk THEN
    bOk := GVL_Devices.aAxis[nAx].bReady AND NOT GVL_Devices.aAxis[nAx].bLockedByKin;
END_IF
IF bOk AND nAx = 1 AND nDir > 0 THEN
    // nicht über die Kollisionsgrenze und nicht in eine Zone mit geschlossenem Niederhalter tippen
    bOk := GVL_Devices.aAxis[1].fActPos < F_Z1Max(GVL_Devices.aAxis[2].fActPos) - 1.0
           AND F_ClampBlocking(GVL_Devices.aAxis[1].fActPos, GVL_Devices.aAxis[1].fActPos + 2.0) = 0;
END_IF
IF bOk AND nAx = 1 AND nDir < 0 THEN
    bOk := F_ClampBlocking(GVL_Devices.aAxis[1].fActPos, GVL_Devices.aAxis[1].fActPos - 2.0) = 0;
END_IF
IF bOk AND nAx >= 1 AND nAx <= 4 THEN
    bOk := (nDir > 0 AND GVL_Devices.aAxis[nAx].fActPos < GVL_Config.aAxisMax[nAx])
        OR (nDir < 0 AND GVL_Devices.aAxis[nAx].fActPos > GVL_Config.aAxisMin[nAx]);
END_IF
IF nJogAxis <> 0 AND (NOT bOk OR nAx <> nJogAxis) THEN
    GVL_Devices.aAxis[nJogAxis].StopJog();
    nJogAxis := 0;
END_IF
IF bOk THEN
    fVel := GVL_Config.aAxisVSetup[nAx] * LIMIT(0.0, GVL_HMI.stCmd.stJog.fVelocityFactor_pct, 100.0) / 100.0
            * GVL_HMI.stStatus.stParamActive.fSingleAxisVelo_pct / 100.0;
    IF fVel > 0.0 THEN
        GVL_Devices.aAxis[nAx].Jog(nDir, fVel);
        nJogAxis := nAx;
    END_IF
END_IF
END_METHOD

END_FUNCTION_BLOCK

// ---- 05_Sequence/FB_ModeManager.TcPOU
// GRAFCET G0 (Not-Halt) und G1 (Betriebsarten) nach [Langfeld].
// 10 Automatik, 11 Pause (Startzustand), 12 Einzelachsen, 13 Rückkehr Grundzustand (ein Zyklus, initialisiert G2/G3).
// Zweistufige Kommandos (S3): erste Stufe und zweite Stufe innerhalb GVL_Config.tTwoStepConfirmation.
FUNCTION_BLOCK FB_ModeManager
VAR_INPUT
    bEStopActive : BOOL;
    bSafetyOk : BOOL;
    nStopCounter : UDINT;       // FB_AlarmManager.nStopCounter: neuer Alarm >= Stop -> Pause
END_VAR
VAR_OUTPUT
    eMode : E_OperatingMode := E_OperatingMode.Pause;
    eG0 : E_G0Step := E_G0Step.S1_Betrieb;
    bFree : BOOL;               // FREI = X10: Abläufe dürfen fahren
    bEnteredPause : BOOL;       // Impuls
    bEnteredSingle : BOOL;      // Impuls: Abläufe abbrechen, Kopplung lösen
    bInitSequences : BOOL;      // Impuls aus Schritt 13: G2 := 20, G3 := 30
    bEnteredAutomatic : BOOL;   // Impuls (Wiederanlauf)
END_VAR
VAR
    nLastStop : UDINT;
    bInit : BOOL := TRUE;
    eFirst : E_HmiCmd := E_HmiCmd.None;
    tFirst : TIME;
    bAckReq : BOOL;
    bSingleReq, bInitReq, bAutoReq, bPauseReq : BOOL;
    eLastMode : E_OperatingMode := E_OperatingMode.Pause;
END_VAR

IF bInit THEN
    nLastStop := nStopCounter;
    bInit := FALSE;
END_IF

// G0 Not-Halt
CASE eG0 OF
E_G0Step.S1_Betrieb:
    IF bEStopActive THEN
        eG0 := E_G0Step.S2_NotHalt;
    END_IF
E_G0Step.S2_NotHalt:
    IF NOT bEStopActive AND bSafetyOk AND bAckReq THEN
        eG0 := E_G0Step.S1_Betrieb;
    END_IF
END_CASE
bAckReq := FALSE;
IF eG0 = E_G0Step.S2_NotHalt AND (eMode = E_OperatingMode.Automatic OR eMode = E_OperatingMode.ReturnToBase) THEN
    eMode := E_OperatingMode.Pause;
END_IF

// Neuer Alarm der Stufe Stop oder Fault -> Pause
IF nStopCounter <> nLastStop THEN
    nLastStop := nStopCounter;
    IF eMode = E_OperatingMode.Automatic OR eMode = E_OperatingMode.ReturnToBase THEN
        eMode := E_OperatingMode.Pause;
    END_IF
END_IF

// Schritt 13: G2/G3 initialisieren, dann Automatik
bInitSequences := bInitReq;
bInitReq := FALSE;
IF eMode = E_OperatingMode.ReturnToBase AND bInitSequences THEN
    eMode := E_OperatingMode.Automatic;
END_IF

bEnteredSingle := bSingleReq;
bSingleReq := FALSE;
bEnteredAutomatic := (eMode = E_OperatingMode.Automatic) AND (eLastMode <> E_OperatingMode.Automatic);
bEnteredPause := (eMode = E_OperatingMode.Pause) AND (eLastMode <> E_OperatingMode.Pause);
eLastMode := eMode;
bFree := eMode = E_OperatingMode.Automatic AND eG0 = E_G0Step.S1_Betrieb;

METHOD CmdPause : E_CmdResult
VAR_INPUT
END_VAR
IF eMode <> E_OperatingMode.Automatic AND eMode <> E_OperatingMode.ReturnToBase THEN
    CmdPause := E_CmdResult.RejectedMode;
    RETURN;
END_IF
eMode := E_OperatingMode.Pause;
CmdPause := E_CmdResult.Accepted;
END_METHOD

METHOD CmdFirstStage : E_CmdResult
// ModeResume1 oder ModeSingleAxis1
VAR_INPUT
    eCmd : E_HmiCmd;
END_VAR
IF eMode <> E_OperatingMode.Pause THEN
    CmdFirstStage := E_CmdResult.RejectedMode;
    RETURN;
END_IF
eFirst := eCmd;
tFirst := TIME();
CmdFirstStage := E_CmdResult.Accepted;
END_METHOD

METHOD CmdSecondStage : E_CmdResult
// ModeResume2 oder ModeSingleAxis2
VAR_INPUT
    eCmd : E_HmiCmd;
    bHmiAlive : BOOL;
    bFaultActive : BOOL;
END_VAR
VAR
    eExpected : E_HmiCmd;
    bOk : BOOL;
END_VAR
IF eMode <> E_OperatingMode.Pause THEN
    CmdSecondStage := E_CmdResult.RejectedMode;
    RETURN;
END_IF
IF eCmd = E_HmiCmd.ModeResume2 THEN
    eExpected := E_HmiCmd.ModeResume1;
ELSE
    eExpected := E_HmiCmd.ModeSingleAxis1;
END_IF
bOk := eFirst = eExpected AND (TIME() - tFirst) <= GVL_Config.tTwoStepConfirmation;
eFirst := E_HmiCmd.None;
IF NOT bOk THEN
    CmdSecondStage := E_CmdResult.RejectedSequence;
    RETURN;
END_IF
IF eCmd = E_HmiCmd.ModeResume2 THEN
    IF NOT bHmiAlive OR eG0 <> E_G0Step.S1_Betrieb OR bFaultActive THEN
        CmdSecondStage := E_CmdResult.RejectedInterlock;
        RETURN;
    END_IF
    eMode := E_OperatingMode.Automatic;
ELSE
    eMode := E_OperatingMode.SingleAxis;
    bSingleReq := TRUE;
END_IF
CmdSecondStage := E_CmdResult.Accepted;
END_METHOD

METHOD CmdReturnToBase : E_CmdResult
VAR_INPUT
    dwMissing : DWORD;      // dwBaseStateMissing
END_VAR
VAR_OUTPUT
    nDetail : UDINT;
END_VAR
IF eMode <> E_OperatingMode.SingleAxis THEN
    CmdReturnToBase := E_CmdResult.RejectedMode;
    RETURN;
END_IF
IF (dwMissing AND 16#3F) <> 0 THEN
    nDetail := DWORD_TO_UDINT(dwMissing AND 16#3F);
    CmdReturnToBase := E_CmdResult.RejectedInterlock;
    RETURN;
END_IF
eMode := E_OperatingMode.ReturnToBase;
bInitReq := TRUE;
CmdReturnToBase := E_CmdResult.Accepted;
END_METHOD

METHOD Acknowledge
// Quittierung (AlarmAck): verlässt G0 Schritt 2, wenn Not-Halt entriegelt und Safety bereit.
VAR_INPUT
END_VAR
bAckReq := TRUE;
END_METHOD

METHOD ForcePause
VAR_INPUT
END_VAR
IF eMode = E_OperatingMode.Automatic OR eMode = E_OperatingMode.ReturnToBase THEN
    eMode := E_OperatingMode.Pause;
END_IF
END_METHOD

END_FUNCTION_BLOCK

// ---- 05_Sequence/FB_BendSequence.TcPOU
// GRAFCET G2 (Biegevorgang, Schritte 20..28) und G3 (Werkstückrotation, 30..32) nach [Langfeld].
// Abweichungen (begründet in docs/grafcet-zuordnung.md):
//  - S21 fährt zusätzlich Z2, X und A an; die Kurvenscheibe des Abschnitts wird in S21 geladen.
//  - Rückbiegen liegt in der Kurvenscheibe (Prüfbericht H4); Geraden zwischen Bögen ohne Halt.
//  - S27 erlaubt nach dem letzten Abschnitt neben ENT auch die Fortsetzung am selben Rohr (Schrittbetrieb).
// Bewegungen nur bei FREI (Automatik). In der Pause hält der Master (Hold) bzw. halten die Einzelbewegungen;
// beim Wiederanlauf setzen die Schritte ihre Bewegungen fort.
FUNCTION_BLOCK FB_BendSequence
VAR_INPUT
    bFree : BOOL;
    bAbort : BOOL;          // Impuls: Wechsel in Einzelachsen -> Ablauf abbrechen
    bInit : BOOL;           // Impuls: G1 Schritt 13 -> G2 := 20, G3 := 30
END_VAR
VAR_OUTPUT
    eStepG2 : E_G2Step := E_G2Step.S20_Grundzustand;
    eStepG3 : E_G3Step := E_G3Step.S30_Bereit;
    nSection : INT;
    bMaterialOk : BOOL;
    bTubeInMachine : BOOL;  // nach dem ersten Start bis ENT
    bWaitingAtEnd : BOOL;   // S27 nach dem letzten Abschnitt: wartet auf ENT oder Fortsetzung
END_VAR
VAR
    ipKin : I_Kinematics;
    eLastG2 : E_G2Step := E_G2Step.S20_Grundzustand;
    bEntry : BOOL;
    bFreeLast : BOOL;
    bQ1, bQ2, bEnt, bContinue : BOOL;
    fWTarget : LREAL;
    tonStep : TON;
    tStepLimit : TIME;
    bOk : BOOL;
    bEndReached : BOOL;
    stKin : ST_KinStatus;
    bAbortReq : BOOL;
    i : INT;
END_VAR

ipKin := GVL_Devices.fbKin;

// ── Abbruch / Initialisierung ──
IF bAbort OR bInit OR bAbortReq THEN
    bAbortReq := FALSE;
    ipKin.Abort();
    FOR i := 1 TO 5 DO
        IF GVL_Devices.aAxis[i].bBusy AND NOT GVL_Devices.aAxis[i].bLockedByKin THEN
            GVL_Devices.aAxis[i].Halt();
        END_IF
    END_FOR
    eStepG2 := E_G2Step.S20_Grundzustand;
    eStepG3 := E_G3Step.S30_Bereit;
    nSection := 0;
    bQ1 := FALSE; bQ2 := FALSE; bEnt := FALSE; bContinue := FALSE;
    IF bInit THEN
        bTubeInMachine := FALSE;
    END_IF
END_IF

// Not-Halt während des Ablaufs: Pneumatik ist entlüftet, die Klemmung nicht mehr gesichert -> Ablauf abbrechen.
// Neustart nur aus der Grundstellung (Prüfbericht: Klemmprüfung nach Not-Halt-Wiederanlauf).
IF GVL_IO.bEStopActive AND eStepG2 <> E_G2Step.S20_Grundzustand AND eStepG2 <> E_G2Step.S27_Uebergabe THEN
    ipKin.Abort();
    eStepG2 := E_G2Step.S20_Grundzustand;
    eStepG3 := E_G3Step.S30_Bereit;
    nSection := 0;
END_IF

// ── Pause und Wiederanlauf ──
IF bFreeLast AND NOT bFree THEN
    ipKin.Hold();
    FOR i := 1 TO 5 DO
        IF GVL_Devices.aAxis[i].bBusy AND NOT GVL_Devices.aAxis[i].bLockedByKin THEN
            GVL_Devices.aAxis[i].Halt();
        END_IF
    END_FOR
ELSIF bFree AND NOT bFreeLast THEN
    IF eStepG2 = E_G2Step.S23_Biegen AND eStepG3 = E_G3Step.S30_Bereit THEN
        ipKin.Resume();
    END_IF
END_IF
bFreeLast := bFree;

bEntry := eStepG2 <> eLastG2;
eLastG2 := eStepG2;

// ── Zeitüberwachung der Bewegungsschritte ──
CASE eStepG2 OF
E_G2Step.S21_Startposition, E_G2Step.S26_Neutral, E_G2Step.S28_Grundstellung:
    tStepLimit := T#120S;
E_G2Step.S22_Niederhalter:
    tStepLimit := T#10S;
ELSE
    tStepLimit := T#0S;
END_CASE
tonStep(IN := bFree AND NOT bEntry AND tStepLimit > T#0S, PT := tStepLimit);
IF tonStep.Q THEN
    GVL_Devices.fbAlarm.Raise(E_AlarmCode.SeqStepTimeout, E_AlarmSeverity.Stop, 0, INT_TO_UDINT(TO_INT(eStepG2)));
    tonStep(IN := FALSE);
END_IF

bWaitingAtEnd := FALSE;

// ── G2 ──
CASE eStepG2 OF
E_G2Step.S20_Grundzustand:
    nSection := 0;

E_G2Step.S21_Startposition:
    IF bEntry THEN
        ipKin.LoadSection(nSection);
    END_IF
    IF bFree THEN
        bOk := MoveTo(2, GVL_Plan.stActive.aSection[nSection].fZ2_mm);
        bOk := MoveTo(3, 0.0) AND bOk;
        bOk := MoveTo(4, 0.0) AND bOk;
        IF bOk THEN   // Z1 erst, wenn Z2 steht (Kollisionsgrenze hängt von Z2 ab)
            IF MoveTo(1, GVL_Plan.stActive.aSection[nSection].fZ1Start_mm) AND ipKin.TableReady() THEN
                eStepG2 := E_G2Step.S22_Niederhalter;
            END_IF
        END_IF
    END_IF

E_G2Step.S22_Niederhalter:
    IF bEntry THEN
        FOR i := 1 TO 6 DO
            IF (GVL_Plan.stActive.aSection[nSection].nClampMask AND SHL(BYTE#1, i - 1)) <> 0
               AND NOT F_ChuckInZone((i + 1) / 2, GVL_Axis.Z1.NcToPlc.ActPos) THEN
                GVL_Devices.aClamp[i].Close();
            END_IF
        END_FOR
    END_IF
    bOk := TRUE;
    FOR i := 1 TO 6 DO
        IF GVL_Devices.aClamp[i].IsCommandedClosed() AND NOT GVL_Devices.aClamp[i].IsClamped() THEN
            bOk := FALSE;
        END_IF
    END_FOR
    IF bOk AND bFree THEN
        eStepG2 := E_G2Step.S23_Biegen;
    END_IF

E_G2Step.S23_Biegen:
    IF bEntry THEN
        ipKin.Start();
    END_IF
    // Niederhalter positionsabhängig öffnen (↑[p_Z1 >= z_NH,i])
    FOR i := 1 TO 6 DO
        IF GVL_Devices.aClamp[i].IsCommandedClosed()
           AND GVL_Axis.Z1.NcToPlc.ActPos >= GVL_Plan.stActive.aSection[nSection].aClampOpen_mm[i] THEN
            GVL_Devices.aClamp[i].Open();
        END_IF
    END_FOR
    IF ipKin.SectionDone() THEN
        eStepG2 := E_G2Step.S24_Halten;
    END_IF

E_G2Step.S24_Halten:
    IF bEntry THEN
        bQ1 := FALSE;
    END_IF
    IF bQ1 THEN
        bQ1 := FALSE;
        eStepG2 := E_G2Step.S25_NhOeffnen;
    END_IF

E_G2Step.S25_NhOeffnen:
    IF bEntry THEN
        bQ2 := FALSE;
        FOR i := 1 TO 6 DO
            GVL_Devices.aClamp[i].Open();
        END_FOR
    END_IF
    IF bQ2 AND AllClampsOpen() THEN
        bQ2 := FALSE;
        eStepG2 := E_G2Step.S26_Neutral;
    END_IF

E_G2Step.S26_Neutral:
    IF bEntry THEN
        ipKin.Abort();
    END_IF
    IF bFree AND NOT ipKin.IsCoupled() THEN
        bOk := MoveTo(3, 0.0);
        bOk := MoveTo(4, 0.0) AND bOk;
        IF bOk THEN
            eStepG2 := E_G2Step.S27_Uebergabe;
        END_IF
    END_IF

E_G2Step.S27_Uebergabe:
    IF bEntry THEN
        nSection := nSection + 1;
        bEnt := FALSE;
        bContinue := FALSE;
        stKin := ipKin.GetStatus();
        bEndReached := NOT GVL_Plan.bValid OR GVL_Plan.stActive.stHeader.nPlanId <> stKin.nPlanId
                       OR nSection > UINT_TO_INT(GVL_Plan.stActive.stHeader.nSectionCount);
    END_IF
    IF NOT bEndReached THEN
        IF bFree THEN
            eStepG2 := E_G2Step.S21_Startposition;
        END_IF
    ELSE
        bWaitingAtEnd := TRUE;
        IF bEnt THEN
            bEnt := FALSE;
            bMaterialOk := FALSE;
            eStepG2 := E_G2Step.S28_Grundstellung;
        ELSIF bContinue THEN
            bContinue := FALSE;
            nSection := 1;
            eStepG2 := E_G2Step.S21_Startposition;
        END_IF
    END_IF

E_G2Step.S28_Grundstellung:
    IF bEntry THEN
        fWTarget := GVL_Devices.aAxis[5].fActPos - F_Mod360(GVL_Devices.aAxis[5].fActPos);
        IF F_Mod360(GVL_Devices.aAxis[5].fActPos) > 180.0 THEN
            fWTarget := fWTarget + 360.0;
        END_IF
    END_IF
    IF bFree THEN
        bOk := MoveTo(2, 0.0);
        bOk := MoveTo(3, 0.0) AND bOk;
        bOk := MoveTo(4, 0.0) AND bOk;
        bOk := MoveTo(5, fWTarget) AND bOk;
        bOk := MoveTo(1, 0.0) AND bOk;
        IF bOk THEN
            bTubeInMachine := FALSE;
            eStepG2 := E_G2Step.S20_Grundzustand;
        END_IF
    END_IF
END_CASE

// ── G3 ──
CASE eStepG3 OF
E_G3Step.S30_Bereit:
    IF eStepG2 = E_G2Step.S23_Biegen AND ipKin.AtRotation() THEN
        eStepG3 := E_G3Step.S31_Stop;
    END_IF

E_G3Step.S31_Stop:
    IF ABS(GVL_Axis.Z1.NcToPlc.ActVelo) < 0.001 THEN
        fWTarget := GVL_Devices.aAxis[5].fActPos + ipKin.RotationAngle();
        eStepG3 := E_G3Step.S32_Drehen;
    END_IF

E_G3Step.S32_Drehen:
    IF bFree AND MoveTo(5, fWTarget) THEN
        IF ipKin.ContinueAfterRotation() THEN
            eStepG3 := E_G3Step.S30_Bereit;
        END_IF
    END_IF
END_CASE

METHOD PRIVATE MoveTo : BOOL
// Fährt Achse nIdx im Eilgang auf fPos, falls sie nicht dort steht. TRUE = angekommen.
VAR_INPUT
    nIdx : INT;
    fPos : LREAL;
END_VAR
IF GVL_Devices.aAxis[nIdx].AtPosition(fPos) THEN
    MoveTo := TRUE;
ELSIF NOT GVL_Devices.aAxis[nIdx].bBusy AND GVL_Devices.aAxis[nIdx].bReady THEN
    GVL_Devices.aAxis[nIdx].MoveAbs(fPos, GVL_Config.aAxisVSetup[nIdx]);
END_IF
END_METHOD

METHOD PRIVATE AllClampsOpen : BOOL
VAR
    k : INT;
END_VAR
AllClampsOpen := TRUE;
FOR k := 1 TO 6 DO
    IF NOT GVL_Devices.aClamp[k].IsOpen() THEN
        AllClampsOpen := FALSE;
    END_IF
END_FOR
END_METHOD

METHOD Start : E_CmdResult
// SeqStart. Betriebsart, Plan, Material, Not-Halt, HMI und Achsen prüft FB_HmiCommand vorher.
// Aus S20 nur in Grundstellung; aus S27 (letzter Abschnitt fertig) als Fortsetzung am selben Rohr.
VAR_INPUT
    dwBaseMissing : DWORD;
END_VAR
VAR_OUTPUT
    nDetail : UDINT;
END_VAR
IF eStepG2 = E_G2Step.S20_Grundzustand THEN
    IF (dwBaseMissing AND 16#3F) <> 0 THEN
        nDetail := DWORD_TO_UDINT(dwBaseMissing AND 16#3F);
        Start := E_CmdResult.RejectedInterlock;
        RETURN;
    END_IF
    nSection := 1;
    bTubeInMachine := TRUE;
    eStepG2 := E_G2Step.S21_Startposition;
    Start := E_CmdResult.Accepted;
ELSIF eStepG2 = E_G2Step.S27_Uebergabe AND bWaitingAtEnd THEN
    IF GVL_Devices.aAxis[1].fActPos > GVL_Plan.stActive.aSection[1].fZ1Start_mm + GVL_Config.fPosTol THEN
        nDetail := 16#20000;
        Start := E_CmdResult.RejectedInterlock;
        RETURN;
    END_IF
    IF (dwBaseMissing AND 16#2C) <> 0 THEN   // X, A nicht auf 0 oder Niederhalter nicht offen
        nDetail := DWORD_TO_UDINT(dwBaseMissing AND 16#2C);
        Start := E_CmdResult.RejectedInterlock;
        RETURN;
    END_IF
    bContinue := TRUE;
    Start := E_CmdResult.Accepted;
ELSE
    Start := E_CmdResult.RejectedSequence;
END_IF
END_METHOD

METHOD ConfirmQ1 : E_CmdResult
VAR_INPUT
END_VAR
IF eStepG2 = E_G2Step.S24_Halten THEN
    bQ1 := TRUE;
    ConfirmQ1 := E_CmdResult.Accepted;
ELSE
    ConfirmQ1 := E_CmdResult.RejectedSequence;
END_IF
END_METHOD

METHOD ConfirmQ2 : E_CmdResult
VAR_INPUT
END_VAR
IF eStepG2 = E_G2Step.S25_NhOeffnen THEN
    bQ2 := TRUE;
    ConfirmQ2 := E_CmdResult.Accepted;
ELSE
    ConfirmQ2 := E_CmdResult.RejectedSequence;
END_IF
END_METHOD

METHOD PartRemoved : E_CmdResult
VAR_INPUT
END_VAR
IF eStepG2 = E_G2Step.S27_Uebergabe AND bWaitingAtEnd THEN
    bEnt := TRUE;
    PartRemoved := E_CmdResult.Accepted;
ELSE
    PartRemoved := E_CmdResult.RejectedSequence;
END_IF
END_METHOD

METHOD CanLoadPlan : BOOL
VAR_INPUT
END_VAR
CanLoadPlan := eStepG2 = E_G2Step.S20_Grundzustand OR (eStepG2 = E_G2Step.S27_Uebergabe AND bWaitingAtEnd);
END_METHOD

METHOD SetMaterial
VAR_INPUT
    bOk : BOOL;
END_VAR
bMaterialOk := bOk;
END_METHOD

METHOD AbortRun
// Ablauf abbrechen (z. B. nach quittiertem Kinematikfehler). Plan bleibt geladen.
VAR_INPUT
END_VAR
bAbortReq := TRUE;
END_METHOD

END_FUNCTION_BLOCK

// ---- 04_Kinematics/F_ChuckInZone.TcPOU
// TRUE, wenn das Futter bei Z1 = fZ1 die Zone des Niederhalterpaares nPair (1..3) berührt.
FUNCTION F_ChuckInZone : BOOL
VAR_INPUT
    nPair : INT;
    fZ1 : LREAL;
END_VAR

IF nPair < 1 OR nPair > 3 THEN
    RETURN;
END_IF
F_ChuckInZone := fZ1 > GVL_Config.aClampZoneLo_mm[nPair] AND fZ1 < GVL_Config.aClampZoneHi_mm[nPair];

END_FUNCTION

// ---- 03_Devices/F_Mod360.TcPOU
// Winkel auf 0 <= Ergebnis < 360 abbilden.
FUNCTION F_Mod360 : LREAL
VAR_INPUT
    fAngle : LREAL;
END_VAR
VAR
    fR : LREAL;
END_VAR

// LREAL_TO_LINT rundet; das Ergebnis liegt dann in [-180, 180] und wird unten korrigiert.
fR := fAngle - 360.0 * LINT_TO_LREAL(LREAL_TO_LINT(fAngle / 360.0));
IF fR < 0.0 THEN
    fR := fR + 360.0;
END_IF
IF fR >= 360.0 THEN
    fR := fR - 360.0;
END_IF
F_Mod360 := fR;

END_FUNCTION

// ---- 06_HMI/FB_PlanStore.TcPOU
// Prüft den Plan im Übergabebereich GVL_HMI.stPlanXfer und übernimmt ihn als aktiven Plan nach GVL_Plan.stActive.
// Rückgabe von Load(): 0 = in Ordnung, sonst Detailcode (backend/biegbert/alarms.py):
//   1 Plan-ID passt nicht, 2 Format/Anzahl/Feld ungültig, 3 Prüfsumme falsch,
//  10 z1_start >= z1_fin, 11 s nicht steigend oder Abschnitte überlappen, 12 u oder phi außerhalb X/A,
//  13 Z2 außerhalb, 14 Ende hinter Kollisionsgrenze, 15 zu viele Punkte, 16 X zu schnell für den Vorschub
FUNCTION_BLOCK FB_PlanStore
VAR
    nLastDetail : UDINT;
END_VAR

;

METHOD Load : UDINT
VAR_INPUT
    nPlanId : UDINT;
END_VAR
VAR
    nSec, nPts, nSc, k, j : INT;
    nFirst, nCnt : INT;
    fPrevFin, fPrevS, fSlope, fFeed, fDs : LREAL;
    nFeedIdx : INT;
END_VAR
Load := 0;
IF nPlanId = 0 OR GVL_HMI.stPlanXfer.stHeader.nPlanId <> nPlanId THEN
    Load := 1; RETURN;
END_IF
IF GVL_HMI.stPlanXfer.stHeader.nFormat <> GVL_Config.cPlanFormat THEN
    Load := 2; RETURN;
END_IF
nSec := UINT_TO_INT(GVL_HMI.stPlanXfer.stHeader.nSectionCount);
IF GVL_HMI.stPlanXfer.stHeader.nPointCount > INT_TO_UDINT(GVL_Config.cMaxPoints) THEN
    Load := 15; RETURN;
END_IF
nPts := UDINT_TO_INT(GVL_HMI.stPlanXfer.stHeader.nPointCount);
IF nSec < 1 OR nSec > GVL_Config.cMaxSections OR nPts < 2 THEN
    Load := 2; RETURN;
END_IF
IF F_PlanChecksum(GVL_HMI.stPlanXfer) <> UDINT_TO_DWORD(GVL_HMI.stPlanXfer.stHeader.nChecksum) THEN
    Load := 3; RETURN;
END_IF

fPrevFin := -1.0E9;
FOR nSc := 1 TO nSec DO
    nFirst := UDINT_TO_INT(GVL_HMI.stPlanXfer.aSection[nSc].nFirstPoint);
    nCnt := UDINT_TO_INT(GVL_HMI.stPlanXfer.aSection[nSc].nPointCount);
    IF NOT (GVL_HMI.stPlanXfer.aSection[nSc].fZ1Start_mm < GVL_HMI.stPlanXfer.aSection[nSc].fZ1Fin_mm) THEN
        Load := 10; RETURN;
    END_IF
    IF nCnt < 2 OR nFirst < 1 OR nFirst + nCnt - 1 > nPts THEN
        Load := 2; RETURN;
    END_IF
    IF GVL_HMI.stPlanXfer.aSection[nSc].fZ1Start_mm < fPrevFin - GVL_Config.fPosTol THEN
        Load := 11; RETURN;
    END_IF
    IF GVL_HMI.stPlanXfer.aSection[nSc].fZ2_mm < GVL_Config.aAxisMin[2] OR GVL_HMI.stPlanXfer.aSection[nSc].fZ2_mm > GVL_Config.aAxisMax[2] THEN
        Load := 13; RETURN;
    END_IF
    IF GVL_HMI.stPlanXfer.aSection[nSc].fZ1Fin_mm > F_Z1Max(GVL_HMI.stPlanXfer.aSection[nSc].fZ2_mm) + GVL_Config.fPosTol
       OR GVL_HMI.stPlanXfer.aSection[nSc].fZ1Fin_mm > GVL_Config.aAxisMax[1] THEN
        Load := 14; RETURN;
    END_IF
    // Vorschubprofil
    IF GVL_HMI.stPlanXfer.aSection[nSc].nFeedCount < 1 OR UINT_TO_INT(GVL_HMI.stPlanXfer.aSection[nSc].nFeedCount) > GVL_Config.cMaxFeed THEN
        Load := 2; RETURN;
    END_IF
    FOR k := 1 TO UINT_TO_INT(GVL_HMI.stPlanXfer.aSection[nSc].nFeedCount) DO
        IF GVL_HMI.stPlanXfer.aSection[nSc].aFeed[k].fFeed_mm_s <= 0.0 OR GVL_HMI.stPlanXfer.aSection[nSc].aFeed[k].fFeed_mm_s > GVL_Config.aAxisVMax[1] THEN
            Load := 2; RETURN;
        END_IF
        IF k > 1 AND_THEN GVL_HMI.stPlanXfer.aSection[nSc].aFeed[k].fZ1_mm <= GVL_HMI.stPlanXfer.aSection[nSc].aFeed[k - 1].fZ1_mm THEN
            Load := 2; RETURN;
        END_IF
    END_FOR
    // Rotationen
    IF UINT_TO_INT(GVL_HMI.stPlanXfer.aSection[nSc].nRotCount) > GVL_Config.cMaxRot THEN
        Load := 2; RETURN;
    END_IF
    FOR k := 1 TO UINT_TO_INT(GVL_HMI.stPlanXfer.aSection[nSc].nRotCount) DO
        IF GVL_HMI.stPlanXfer.aSection[nSc].aRot[k].fZ1_mm < GVL_HMI.stPlanXfer.aSection[nSc].fZ1Start_mm - GVL_Config.fPosTol
           OR GVL_HMI.stPlanXfer.aSection[nSc].aRot[k].fZ1_mm > GVL_HMI.stPlanXfer.aSection[nSc].fZ1Fin_mm + GVL_Config.fPosTol
           OR (k > 1 AND_THEN GVL_HMI.stPlanXfer.aSection[nSc].aRot[k].fZ1_mm < GVL_HMI.stPlanXfer.aSection[nSc].aRot[k - 1].fZ1_mm) THEN
            Load := 2; RETURN;
        END_IF
    END_FOR
    // Stützpunkte
    IF ABS(GVL_HMI.stPlanXfer.aPoint[nFirst].fS_mm - GVL_HMI.stPlanXfer.aSection[nSc].fZ1Start_mm) > GVL_Config.fPosTol
       OR ABS(GVL_HMI.stPlanXfer.aPoint[nFirst + nCnt - 1].fS_mm - GVL_HMI.stPlanXfer.aSection[nSc].fZ1Fin_mm) > GVL_Config.fPosTol THEN
        Load := 11; RETURN;
    END_IF
    nFeedIdx := 1;
    FOR j := nFirst TO nFirst + nCnt - 1 DO
        IF ABS(GVL_HMI.stPlanXfer.aPoint[j].fU_mm) > GVL_Config.aAxisMax[3] OR ABS(GVL_HMI.stPlanXfer.aPoint[j].fPhi_deg) > GVL_Config.aAxisMax[4] THEN
            Load := 12; RETURN;
        END_IF
        IF j > nFirst THEN
            fDs := GVL_HMI.stPlanXfer.aPoint[j].fS_mm - GVL_HMI.stPlanXfer.aPoint[j - 1].fS_mm;
            IF fDs <= 0.0 THEN
                Load := 11; RETURN;
            END_IF
            WHILE nFeedIdx < UINT_TO_INT(GVL_HMI.stPlanXfer.aSection[nSc].nFeedCount)
                  AND_THEN GVL_HMI.stPlanXfer.aSection[nSc].aFeed[nFeedIdx + 1].fZ1_mm <= GVL_HMI.stPlanXfer.aPoint[j - 1].fS_mm + 1.0E-6 DO
                nFeedIdx := nFeedIdx + 1;
            END_WHILE
            fFeed := GVL_HMI.stPlanXfer.aSection[nSc].aFeed[nFeedIdx].fFeed_mm_s;
            fSlope := ABS(GVL_HMI.stPlanXfer.aPoint[j].fU_mm - GVL_HMI.stPlanXfer.aPoint[j - 1].fU_mm) / fDs;
            IF fSlope * fFeed > GVL_Config.aAxisVMax[3] * 1.05 THEN
                Load := 16; RETURN;
            END_IF
        END_IF
    END_FOR
    fPrevFin := GVL_HMI.stPlanXfer.aSection[nSc].fZ1Fin_mm;
END_FOR

MEMCPY(destAddr := ADR(GVL_Plan.stActive), srcAddr := ADR(GVL_HMI.stPlanXfer), n := SIZEOF(ST_PlanTransfer));
GVL_Plan.bValid := TRUE;
END_METHOD

METHOD Invalidate
VAR_INPUT
END_VAR
GVL_Plan.bValid := FALSE;
GVL_Plan.stActive.stHeader.nPlanId := 0;
END_METHOD

END_FUNCTION_BLOCK

// ---- 06_HMI/F_PlanChecksum.TcPOU
// Prüfsumme über die belegten Abschnitte und Punkte eines Plans (gleicher Algorithmus in backend/biegbert/plc/layout.py):
// h := ROL(h, 5) XOR Byte, Startwert 0.
FUNCTION F_PlanChecksum : DWORD
VAR_IN_OUT
    stPlan : ST_PlanTransfer;
END_VAR
VAR
    p : POINTER TO BYTE;
    n, i : UDINT;
    h : DWORD;
END_VAR

h := 0;
p := ADR(stPlan.aSection[1]);
n := UINT_TO_UDINT(stPlan.stHeader.nSectionCount) * SIZEOF(ST_PlanSection);
FOR i := 1 TO n DO
    h := ROL(h, 5) XOR BYTE_TO_DWORD(p^);
    p := p + 1;
END_FOR
p := ADR(stPlan.aPoint[1]);
n := stPlan.stHeader.nPointCount * SIZEOF(ST_PlanPoint);
FOR i := 1 TO n DO
    h := ROL(h, 5) XOR BYTE_TO_DWORD(p^);
    p := p + 1;
END_FOR
F_PlanChecksum := h;

END_FUNCTION

// ---- 04_Kinematics/F_Z1Max.TcPOU
// Größte zulässige Z1-Position (Futter <-> Führung) bei gegebener Z2-Position.
FUNCTION F_Z1Max : LREAL
VAR_INPUT
    fZ2 : LREAL;
END_VAR

F_Z1Max := GVL_Config.fZ1CollisionBase_mm + fZ2;

END_FUNCTION

// ---- 04_Kinematics/F_ClampBlocking.TcPOU
// Paar (1..3), dessen Zone eine Z1-Fahrt von fFrom nach fTo kreuzt, obwohl einer seiner Niederhalter nicht offen ist; 0 = frei.
FUNCTION F_ClampBlocking : INT
VAR_INPUT
    fFrom : LREAL;
    fTo : LREAL;
END_VAR
VAR
    p : INT;
    a, b : LREAL;
END_VAR

a := MIN(fFrom, fTo);
b := MAX(fFrom, fTo);
FOR p := 1 TO 3 DO
    IF b > GVL_Config.aClampZoneLo_mm[p] AND a < GVL_Config.aClampZoneHi_mm[p] THEN
        IF NOT GVL_Devices.aClamp[2 * p - 1].IsOpen() OR NOT GVL_Devices.aClamp[2 * p].IsOpen() THEN
            F_ClampBlocking := p;
            RETURN;
        END_IF
    END_IF
END_FOR

END_FUNCTION

// ---- 05_Sequence/FB_Interlocks.TcPOU
// Zyklische Überwachung über mehrere Geräte: Abstand Futter <-> Führung, Futter in Niederhalterzone,
// Software-Endlagen, Achs- und Niederhalterfehler, Not-Halt. Setzt und löscht die zugehörigen Alarme.
FUNCTION_BLOCK FB_Interlocks
VAR
    i, p, k : INT;
    fZ1, fZmax : LREAL;
    bViolation : BOOL;
    bOut : BOOL;
END_VAR

fZ1 := GVL_Devices.aAxis[1].fActPos;
fZmax := F_Z1Max(GVL_Devices.aAxis[2].fActPos);

// Abstand Futter <-> Führung (dZ12)
IF fZ1 > fZmax + GVL_Config.fPosTol THEN
    IF NOT GVL_Devices.fbAlarm.IsActive(E_AlarmCode.DistanceZ1Z2, 1, FALSE) THEN
        StopZ1();
        GVL_Devices.fbAlarm.Raise(E_AlarmCode.DistanceZ1Z2, E_AlarmSeverity.Stop, 1, 0);
    END_IF
ELSIF fZ1 < fZmax - 1.0 THEN
    GVL_Devices.fbAlarm.Clear(E_AlarmCode.DistanceZ1Z2, 1, FALSE);
END_IF

// Futter in der Zone eines nicht offenen Niederhalters
FOR p := 1 TO 3 DO
    FOR k := 2 * p - 1 TO 2 * p DO
        bViolation := F_ChuckInZone(p, fZ1)
                      AND (GVL_Devices.aClamp[k].IsCommandedClosed() OR GVL_Devices.aClamp[k].eState = E_ClampState.Closing
                           OR GVL_Devices.aClamp[k].eState = E_ClampState.Clamped);
        IF bViolation AND NOT GVL_Devices.fbAlarm.IsActive(E_AlarmCode.ClampZoneViolation, k, FALSE) THEN
            StopZ1();
            GVL_Devices.fbAlarm.Raise(E_AlarmCode.ClampZoneViolation, E_AlarmSeverity.Fault, k, 0);
        ELSIF NOT bViolation THEN
            GVL_Devices.fbAlarm.Clear(E_AlarmCode.ClampZoneViolation, k, FALSE);
        END_IF
    END_FOR
END_FOR

// Achsen: Fehler und Software-Endlagen (W ist endlos)
FOR i := 1 TO 5 DO
    GVL_Devices.fbAlarm.Set(GVL_Devices.aAxis[i].bError, E_AlarmCode.AxisError, E_AlarmSeverity.Fault, i,
                            GVL_Devices.aAxis[i].nErrorId);
    IF i < 5 THEN
        bOut := GVL_Devices.aAxis[i].fActPos > GVL_Config.aAxisMax[i] + GVL_Config.fPosTol
             OR GVL_Devices.aAxis[i].fActPos < GVL_Config.aAxisMin[i] - GVL_Config.fPosTol;
        IF bOut AND NOT GVL_Devices.fbAlarm.IsActive(E_AlarmCode.AxisSoftLimit, i, FALSE) THEN
            IF GVL_Devices.aAxis[i].IsJogging() THEN
                GVL_Devices.aAxis[i].StopJog();
            END_IF
        END_IF
        GVL_Devices.fbAlarm.Set(bOut, E_AlarmCode.AxisSoftLimit, E_AlarmSeverity.Warning, i, 0);
    END_IF
END_FOR

// Niederhalter
FOR k := 1 TO 6 DO
    GVL_Devices.fbAlarm.Set(GVL_Devices.aClamp[k].bTimeoutFault, E_AlarmCode.ClampTimeout, E_AlarmSeverity.Fault, k, 0);
    GVL_Devices.fbAlarm.Set(GVL_Devices.aClamp[k].bPressureFault, E_AlarmCode.ClampPressureLow, E_AlarmSeverity.Fault, k, 0);
END_FOR

// Not-Halt und Safety
GVL_Devices.fbAlarm.Set(GVL_IO.bEStopActive, E_AlarmCode.EStopActive, E_AlarmSeverity.Fault, 0, 0);
GVL_Devices.fbAlarm.Set(NOT GVL_IO.bSafetyOk, E_AlarmCode.SafetyNotReady, E_AlarmSeverity.Fault, 0, 0);

METHOD PRIVATE StopZ1
VAR_INPUT
END_VAR
IF GVL_Devices.fbKin.IsCoupled() THEN
    GVL_Devices.fbKin.Hold();
ELSE
    GVL_Devices.aAxis[1].Halt();
END_IF
END_METHOD

END_FUNCTION_BLOCK

// ---- 06_HMI/FB_HmiStatus.TcPOU
// Füllt GVL_HMI.stStatus (stCmdAck und stParamActive pflegt FB_HmiCommand).
FUNCTION_BLOCK FB_HmiStatus
VAR_IN_OUT
    fbMode : FB_ModeManager;
    fbSeq : FB_BendSequence;
END_VAR
VAR_INPUT
    bHmiAlive : BOOL;
    bSimulation : BOOL;
    dwBaseMissing : DWORD;
END_VAR
VAR
    i : INT;
END_VAR

GVL_HMI.stStatus.nLifeCounter := GVL_HMI.stStatus.nLifeCounter + 1;
GVL_HMI.stStatus.bHmiAlive := bHmiAlive;
GVL_HMI.stStatus.bSimulation := bSimulation;
GVL_HMI.stStatus.bEStopActive := GVL_IO.bEStopActive;
GVL_HMI.stStatus.bSafetyOk := GVL_IO.bSafetyOk;
GVL_HMI.stStatus.eMode := fbMode.eMode;
GVL_HMI.stStatus.nStepG2 := TO_INT(fbSeq.eStepG2);
GVL_HMI.stStatus.nStepG3 := TO_INT(fbSeq.eStepG3);
GVL_HMI.stStatus.nBend := INT_TO_UDINT(MAX(0, fbSeq.nSection));
GVL_HMI.stStatus.dwBaseStateMissing := dwBaseMissing;

FOR i := 1 TO 5 DO
    GVL_HMI.stStatus.aAxis[i].eState := GVL_Devices.aAxis[i].eState;
    GVL_HMI.stStatus.aAxis[i].bEnabled := GVL_Devices.aAxis[i].bEnabled;
    GVL_HMI.stStatus.aAxis[i].bReady := GVL_Devices.aAxis[i].bReady;
    GVL_HMI.stStatus.aAxis[i].bError := GVL_Devices.aAxis[i].bError;
    GVL_HMI.stStatus.aAxis[i].nErrorId := GVL_Devices.aAxis[i].nErrorId;
    IF i = 5 THEN
        GVL_HMI.stStatus.aAxis[i].fActPos := F_Mod360(GVL_Devices.aAxis[i].fActPos);
        GVL_HMI.stStatus.aAxis[i].fSetPos := F_Mod360(GVL_Devices.aAxis[i].fSetPos);
    ELSE
        GVL_HMI.stStatus.aAxis[i].fActPos := GVL_Devices.aAxis[i].fActPos;
        GVL_HMI.stStatus.aAxis[i].fSetPos := GVL_Devices.aAxis[i].fSetPos;
    END_IF
    GVL_HMI.stStatus.aAxis[i].fActVelo := GVL_Devices.aAxis[i].fActVelo;
    GVL_HMI.stStatus.aAxis[i].fSetVelo := GVL_Devices.aAxis[i].fSetVelo;
    GVL_HMI.stStatus.aAxis[i].fLagError := GVL_Devices.aAxis[i].fLag;
    GVL_HMI.stStatus.aAxis[i].fTorque_Nm := GVL_IO.afTorque_Nm[i];
END_FOR
FOR i := 1 TO 6 DO
    GVL_HMI.stStatus.aClamp[i].eState := GVL_Devices.aClamp[i].eState;
    GVL_HMI.stStatus.aClamp[i].bValve := GVL_Devices.aClamp[i].bValve;
    GVL_HMI.stStatus.aClamp[i].bOpen := GVL_IO.abClampOpen[i];
    GVL_HMI.stStatus.aClamp[i].fLastSwitchTime_ms := GVL_Devices.aClamp[i].fLastSwitchTime_ms;
END_FOR
GVL_HMI.stStatus.stIo.bPressureOk := GVL_IO.bPressureOk;
GVL_HMI.stStatus.stIo.abPanelIn := GVL_IO.abPanel;
GVL_HMI.stStatus.stIo.abPanelOut := GVL_IO.abPanelLamp;
GVL_HMI.stStatus.stKin := GVL_Devices.fbKin.GetStatus();

METHOD CalcBaseMissing : DWORD
// Fehlende Grundzustandsbedingungen (Bits wie docs/hmi-schnittstelle.md).
VAR_INPUT
    bMaterialOk : BOOL;
END_VAR
VAR
    dw : DWORD;
    k : INT;
    fPos : LREAL;
    stKin : ST_KinStatus;
END_VAR
dw := 0;
FOR k := 1 TO 5 DO
    fPos := GVL_Devices.aAxis[k].fActPos;
    IF k = 5 THEN
        fPos := F_Mod360(fPos + 180.0) - 180.0;
    END_IF
    IF ABS(fPos) > GVL_Config.fPosTol THEN
        dw := dw OR SHL(DWORD#1, k - 1);
    END_IF
END_FOR
FOR k := 1 TO 6 DO
    IF NOT GVL_Devices.aClamp[k].IsOpen() THEN
        dw := dw OR 16#20;
    END_IF
END_FOR
IF GVL_Devices.fbAlarm.FaultActive() THEN
    dw := dw OR 16#40;
END_IF
FOR k := 1 TO 5 DO
    IF GVL_Devices.aAxis[k].bError THEN
        dw := dw OR 16#40;
    END_IF
END_FOR
IF NOT GVL_IO.bSafetyOk THEN
    dw := dw OR 16#80;
END_IF
stKin := GVL_Devices.fbKin.GetStatus();
IF stKin.nPlanId = 0 OR NOT GVL_Plan.bValid THEN
    dw := dw OR 16#100;
END_IF
IF NOT bMaterialOk THEN
    dw := dw OR 16#200;
END_IF
CalcBaseMissing := dw;
END_METHOD

END_FUNCTION_BLOCK

// ---- 07_Test/PRG_TEST.TcPOU
PROGRAM PRG_TEST
VAR
    fbBendKinematics_Test : FB_BendKinematics_Test;
END_VAR

TcUnit.RUN();

END_PROGRAM

// ---- 07_Test/FB_BendKinematics_Test.TcPOU
// TcUnit-Tests ohne Achsen: Kinematik-Zustände ohne Plan, Alarmverwaltung, Niederhalter-Zustandsautomat.
// Läuft nur mit Compiler-Define TEST (MAIN ruft PRG_TEST).
FUNCTION_BLOCK FB_BendKinematics_Test EXTENDS TcUnit.FB_TestSuite
VAR
END_VAR

StartWithoutPlanIsRejected();
LoadPlanWithoutValidPlanIsRejected();
AlarmIsRemovedAfterClearAndAck();
StopAlarmCountsStopEvent();

METHOD StartWithoutPlanIsRejected
VAR
    fbKin : FB_BendKinematics;
END_VAR
TEST('StartWithoutPlanIsRejected');
AssertFalse(Condition := fbKin.Start(), Message := 'Start ohne Plan muss abgelehnt werden');
TEST_FINISHED();
END_METHOD

METHOD LoadPlanWithoutValidPlanIsRejected
VAR
    fbKin : FB_BendKinematics;
END_VAR
TEST('LoadPlanWithoutValidPlanIsRejected');
GVL_Plan.bValid := FALSE;
AssertFalse(Condition := fbKin.LoadPlan(nPlanId := 7), Message := 'LoadPlan ohne geprüften Plan muss abgelehnt werden');
TEST_FINISHED();
END_METHOD

METHOD AlarmIsRemovedAfterClearAndAck
VAR
    fbAl : FB_AlarmManager;
    stOut : ST_HmiAlarms;
END_VAR
TEST('AlarmIsRemovedAfterClearAndAck');
fbAl.Raise(E_AlarmCode.ClampTimeout, E_AlarmSeverity.Fault, 3, 0);
fbAl.WriteTo(stOut);
AssertEquals_UINT(Expected := 1, Actual := stOut.nCount, Message := 'ein Eintrag erwartet');
AssertTrue(Condition := fbAl.FaultActive(), Message := 'Fault muss aktiv sein');
fbAl.Ack(0);
fbAl.WriteTo(stOut);
AssertEquals_UINT(Expected := 1, Actual := stOut.nCount, Message := 'quittiert, aber Ursache besteht noch');
fbAl.Clear(E_AlarmCode.ClampTimeout, 3, FALSE);
fbAl.WriteTo(stOut);
AssertEquals_UINT(Expected := 0, Actual := stOut.nCount, Message := 'Eintrag muss entfernt sein');
TEST_FINISHED();
END_METHOD

METHOD StopAlarmCountsStopEvent
VAR
    fbAl : FB_AlarmManager;
END_VAR
TEST('StopAlarmCountsStopEvent');
fbAl.Raise(E_AlarmCode.AxisSoftLimit, E_AlarmSeverity.Warning, 1, 0);
AssertEquals_UDINT(Expected := 0, Actual := fbAl.nStopCounter, Message := 'Warnung darf nicht pausieren');
fbAl.Raise(E_AlarmCode.HmiHeartbeatLost, E_AlarmSeverity.Stop, 0, 0);
AssertEquals_UDINT(Expected := 1, Actual := fbAl.nStopCounter, Message := 'Stop muss zählen');
TEST_FINISHED();
END_METHOD

END_FUNCTION_BLOCK

// ---- 04_Kinematics/FB_BendKinematics.TcPOU
// Kopplung Z1 (Master) -> X, A (Slaves) mit NC Camming (E6). Eine Kurvenscheibe je Planabschnitt; Geraden sind
// Teil der Kurvenscheibe (u = 0), dadurch kein Halt zwischen Bögen. Der Master hält nur an Rotationen (G3) und am
// Abschnittsende. Vorschub stückweise nach dem Vorschubprofil des Abschnitts. Zustände: docs/kinematik.md
FUNCTION_BLOCK FB_BendKinematics IMPLEMENTS I_Kinematics
VAR
    stStatus : ST_KinStatus := (eMode := E_MotionMode.Single);
    nSection : INT;
    bTableReady : BOOL;
    bLoading : BOOL;
    bAtRot : BOOL;
    bDone : BOOL;
    nRotIdx : INT;            // nächste offene Rotation im Abschnitt
    fTargetCmd : LREAL;
    fFeedCmd : LREAL;
    bMasterActive : BOOL;
    bMasterReq : BOOL;
    bHaltActive : BOOL;
    nPhase : INT;             // Unterschritte in Coupling, Decoupling, Fault

    aCamX : ARRAY[1..4000, 1..2] OF LREAL;   // Spalte 1 = Z1, Spalte 2 = X
    aCamA : ARRAY[1..4000, 1..2] OF LREAL;   // Spalte 1 = Z1, Spalte 2 = A
    stCamX : MC_CAM_REF;
    stCamA : MC_CAM_REF;
    fbSelX : MC_CamTableSelect;
    fbSelA : MC_CamTableSelect;
    fbInX : MC_CamIn;
    fbInA : MC_CamIn;
    fbOutX : MC_CamOut;
    fbOutA : MC_CamOut;
    fbMaster : MC_MoveAbsolute;
    fbHalt : MC_Halt;
    bSelExec, bInExec, bOutExec : BOOL;
    bHoldPending : BOOL;      // Hold() während Coupling: nach dem Koppeln nicht losfahren
END_VAR
VAR CONSTANT
    cTableX : UDINT := 1;
    cTableA : UDINT := 2;
END_VAR

// Aufruf über Cyclic().

METHOD Cyclic
VAR_INPUT
END_VAR
VAR
    fZ1 : LREAL;
    fFeed : LREAL;
    fTarget : LREAL;
    nErr : UDINT;
END_VAR
fZ1 := GVL_Axis.Z1.NcToPlc.ActPos;
stStatus.fMasterPos_mm := fZ1;

// ── Kurvenscheiben laden ──
fbSelX(Master := GVL_Axis.Z1, Slave := GVL_Axis.X, CamTable := stCamX, Execute := bSelExec,
       Periodic := FALSE, MasterAbsolute := TRUE, SlaveAbsolute := TRUE, CamTableID := cTableX);
fbSelA(Master := GVL_Axis.Z1, Slave := GVL_Axis.A, CamTable := stCamA, Execute := bSelExec,
       Periodic := FALSE, MasterAbsolute := TRUE, SlaveAbsolute := TRUE, CamTableID := cTableA);
IF bLoading THEN
    IF fbSelX.Error OR fbSelA.Error THEN
        bLoading := FALSE;
        bSelExec := FALSE;
        IF fbSelX.Error THEN nErr := fbSelX.ErrorID; ELSE nErr := fbSelA.ErrorID; END_IF
        GVL_Devices.fbAlarm.Raise(E_AlarmCode.KinCoupleFailed, E_AlarmSeverity.Fault, 0, nErr);
        stStatus.eState := E_KinState.Fault;
        stStatus.nErrorId := nErr;
    ELSIF fbSelX.Done AND fbSelA.Done THEN
        bLoading := FALSE;
        bSelExec := FALSE;
        bTableReady := TRUE;
    END_IF
END_IF

// ── Kopplung ──
fbInX(Master := GVL_Axis.Z1, Slave := GVL_Axis.X, Execute := bInExec, MasterOffset := 0.0, SlaveOffset := 0.0,
      MasterScaling := 1.0, SlaveScaling := 1.0, StartMode := MC_StartMode.MC_STARTMODE_ABSOLUTE, CamTableID := cTableX);
fbInA(Master := GVL_Axis.Z1, Slave := GVL_Axis.A, Execute := bInExec, MasterOffset := 0.0, SlaveOffset := 0.0,
      MasterScaling := 1.0, SlaveScaling := 1.0, StartMode := MC_StartMode.MC_STARTMODE_ABSOLUTE, CamTableID := cTableA);
fbOutX(Slave := GVL_Axis.X, Execute := bOutExec);
fbOutA(Slave := GVL_Axis.A, Execute := bOutExec);

// ── Master: Fahrauftrag und Halt ──
IF bMasterReq THEN
    bMasterReq := FALSE;
    fbMaster(Axis := GVL_Axis.Z1, Execute := FALSE);
    bMasterActive := TRUE;
END_IF
fbMaster(Axis := GVL_Axis.Z1, Execute := bMasterActive, Position := fTargetCmd, Velocity := fFeedCmd,
         Acceleration := GVL_Config.aAxisAccel[1], Deceleration := GVL_Config.aAxisAccel[1]);
fbHalt(Axis := GVL_Axis.Z1, Execute := bHaltActive, Deceleration := GVL_Config.aAxisAccel[1]);

// ── Überwachung im gekoppelten Betrieb ──
CASE stStatus.eState OF
E_KinState.Coupling, E_KinState.Running, E_KinState.Holding, E_KinState.Held:
    IF GVL_Devices.aAxis[1].bError THEN
        EnterFault(E_AlarmCode.KinMasterFault, GVL_Devices.aAxis[1].nErrorId);
    ELSIF GVL_Devices.aAxis[3].bError THEN
        EnterFault(E_AlarmCode.KinSlaveFault, GVL_Devices.aAxis[3].nErrorId);
    ELSIF GVL_Devices.aAxis[4].bError THEN
        EnterFault(E_AlarmCode.KinSlaveFault, GVL_Devices.aAxis[4].nErrorId);
    ELSIF fbInX.Error OR fbInA.Error THEN
        IF fbInX.Error THEN nErr := fbInX.ErrorID; ELSE nErr := fbInA.ErrorID; END_IF
        EnterFault(E_AlarmCode.KinCoupleFailed, nErr);
    ELSIF fbMaster.Error THEN
        EnterFault(E_AlarmCode.KinMasterFault, fbMaster.ErrorID);
    END_IF
END_CASE

// ── Zustände ──
CASE stStatus.eState OF
E_KinState.Coupling:
    bInExec := TRUE;
    IF fbInX.InSync AND fbInA.InSync THEN
        IF bHoldPending THEN
            bHoldPending := FALSE;
            stStatus.eState := E_KinState.Held;
        ELSE
            stStatus.eState := E_KinState.Running;
            IssueMaster(TRUE);
        END_IF
    END_IF

E_KinState.Running:
    fFeed := DesiredFeed(fZ1);
    fTarget := NextStop();
    IF ABS(fFeed - fFeedCmd) > 1.0E-6 OR ABS(fTarget - fTargetCmd) > 1.0E-6 THEN
        IssueMaster(FALSE);
    END_IF
    IF bMasterActive AND fbMaster.Done THEN
        bMasterActive := FALSE;
        IF ABS(fZ1 - GVL_Plan.stActive.aSection[nSection].fZ1Fin_mm) <= GVL_Config.fPosTol
           AND nRotIdx > UINT_TO_INT(GVL_Plan.stActive.aSection[nSection].nRotCount) THEN
            bDone := TRUE;
        ELSE
            bAtRot := TRUE;
        END_IF
        stStatus.eState := E_KinState.Held;
    END_IF

E_KinState.Holding:
    IF NOT bHaltActive THEN
        bMasterActive := FALSE;
        fbHalt(Axis := GVL_Axis.Z1, Execute := FALSE);
        bHaltActive := TRUE;
    ELSIF fbHalt.Done OR fbHalt.Error OR fbHalt.CommandAborted THEN
        bHaltActive := FALSE;
        stStatus.eState := E_KinState.Held;
    END_IF

E_KinState.Decoupling:
    CASE nPhase OF
    0:  // Master anhalten
        bMasterActive := FALSE;
        IF ABS(GVL_Axis.Z1.NcToPlc.ActVelo) > 0.001 THEN
            fbHalt(Axis := GVL_Axis.Z1, Execute := FALSE);
            bHaltActive := TRUE;
            nPhase := 1;
        ELSE
            nPhase := 2;
        END_IF
    1:
        IF fbHalt.Done OR fbHalt.Error OR fbHalt.CommandAborted THEN
            bHaltActive := FALSE;
            nPhase := 2;
        END_IF
    2:  // Slaves auskoppeln (erst im Stillstand des Masters)
        bInExec := FALSE;
        bOutExec := TRUE;
        nPhase := 3;
    3:
        IF (fbOutX.Done OR fbOutX.Error) AND (fbOutA.Done OR fbOutA.Error) THEN
            bOutExec := FALSE;
            nPhase := 0;
            bTableReady := FALSE;
            bAtRot := FALSE;
            bDone := FALSE;
            IF GVL_Plan.bValid AND stStatus.nPlanId <> 0 THEN
                stStatus.eState := E_KinState.Loaded;
            ELSE
                stStatus.eState := E_KinState.Idle;
            END_IF
        END_IF
    END_CASE

E_KinState.Fault:
    // Master stoppen, dann Slaves auskoppeln; bleibt Fault bis Reset()
    CASE nPhase OF
    0:
        bMasterActive := FALSE;
        IF NOT GVL_Devices.aAxis[1].bError AND ABS(GVL_Axis.Z1.NcToPlc.ActVelo) > 0.001 THEN
            fbHalt(Axis := GVL_Axis.Z1, Execute := FALSE);
            bHaltActive := TRUE;
        END_IF
        nPhase := 1;
    1:
        IF NOT bHaltActive OR fbHalt.Done OR fbHalt.Error OR fbHalt.CommandAborted THEN
            bHaltActive := FALSE;
            bInExec := FALSE;
            bOutExec := TRUE;
            nPhase := 2;
        END_IF
    2:
        IF (fbOutX.Done OR fbOutX.Error) AND (fbOutA.Done OR fbOutA.Error) THEN
            bOutExec := FALSE;
            nPhase := 3;
        END_IF
    END_CASE
END_CASE

CASE stStatus.eState OF
E_KinState.Coupling, E_KinState.Running:
    stStatus.eMode := E_MotionMode.Coupled;
E_KinState.Holding, E_KinState.Held:
    stStatus.eMode := E_MotionMode.Hold;
ELSE
    stStatus.eMode := E_MotionMode.Single;
END_CASE
stStatus.bError := stStatus.eState = E_KinState.Fault;
END_METHOD

METHOD PRIVATE EnterFault
VAR_INPUT
    eCode : E_AlarmCode;
    nErr : UDINT;
END_VAR
GVL_Devices.fbAlarm.Raise(eCode, E_AlarmSeverity.Fault, 0, nErr);
stStatus.nErrorId := nErr;
stStatus.eState := E_KinState.Fault;
bHaltActive := FALSE;
nPhase := 0;
END_METHOD

METHOD PRIVATE FeedAt : LREAL
VAR_INPUT
    fZ1 : LREAL;
END_VAR
VAR
    k : INT;
END_VAR
FeedAt := GVL_Plan.stActive.aSection[nSection].aFeed[1].fFeed_mm_s;
FOR k := 2 TO UINT_TO_INT(GVL_Plan.stActive.aSection[nSection].nFeedCount) DO
    IF fZ1 >= GVL_Plan.stActive.aSection[nSection].aFeed[k].fZ1_mm - 1.0E-6 THEN
        FeedAt := GVL_Plan.stActive.aSection[nSection].aFeed[k].fFeed_mm_s;
    END_IF
END_FOR
END_METHOD

METHOD PRIVATE DesiredFeed : LREAL
// Vorschub mit Vorausschau um den Bremsweg: vor einer Biegezone schon langsam sein, damit X nicht überfordert wird.
VAR_INPUT
    fZ1 : LREAL;
END_VAR
VAR
    v0 : LREAL;
END_VAR
v0 := MAX(fFeedCmd, FeedAt(fZ1));
DesiredFeed := FeedAhead(fZ1, v0 * v0 / (2.0 * GVL_Config.aAxisAccel[1]) + 1.0);
END_METHOD

METHOD PRIVATE FeedAhead : LREAL
// Kleinster Vorschub im Bereich [fZ1, fZ1 + fLook].
VAR_INPUT
    fZ1 : LREAL;
    fLook : LREAL;
END_VAR
VAR
    k : INT;
END_VAR
FeedAhead := FeedAt(fZ1);
FOR k := 1 TO UINT_TO_INT(GVL_Plan.stActive.aSection[nSection].nFeedCount) DO
    IF GVL_Plan.stActive.aSection[nSection].aFeed[k].fZ1_mm > fZ1
       AND GVL_Plan.stActive.aSection[nSection].aFeed[k].fZ1_mm <= fZ1 + fLook THEN
        FeedAhead := MIN(FeedAhead, GVL_Plan.stActive.aSection[nSection].aFeed[k].fFeed_mm_s);
    END_IF
END_FOR
END_METHOD

METHOD PRIVATE NextStop : LREAL
VAR_INPUT
END_VAR
IF nRotIdx <= UINT_TO_INT(GVL_Plan.stActive.aSection[nSection].nRotCount) THEN
    NextStop := GVL_Plan.stActive.aSection[nSection].aRot[nRotIdx].fZ1_mm;
ELSE
    NextStop := GVL_Plan.stActive.aSection[nSection].fZ1Fin_mm;
END_IF
END_METHOD

METHOD PRIVATE IssueMaster
VAR_INPUT
    bForce : BOOL;
END_VAR
fFeedCmd := DesiredFeed(GVL_Axis.Z1.NcToPlc.ActPos);
fTargetCmd := NextStop();
bMasterReq := TRUE;
END_METHOD

METHOD LoadPlan : BOOL
VAR_INPUT
    nPlanId : UDINT;
END_VAR
IF (stStatus.eState = E_KinState.Idle OR stStatus.eState = E_KinState.Loaded)
   AND GVL_Plan.bValid AND GVL_Plan.stActive.stHeader.nPlanId = nPlanId AND nPlanId <> 0 THEN
    stStatus.nPlanId := nPlanId;
    stStatus.eState := E_KinState.Loaded;
    nSection := 0;
    bTableReady := FALSE;
    LoadPlan := TRUE;
END_IF
END_METHOD

METHOD LoadSection : BOOL
VAR_INPUT
    nSection : INT;
END_VAR
VAR
    i, n, nFirst : INT;
END_VAR
IF stStatus.eState <> E_KinState.Loaded OR bLoading OR NOT GVL_Plan.bValid
   OR nSection < 1 OR nSection > UINT_TO_INT(GVL_Plan.stActive.stHeader.nSectionCount) THEN
    RETURN;
END_IF
THIS^.nSection := nSection;
nFirst := UDINT_TO_INT(GVL_Plan.stActive.aSection[nSection].nFirstPoint);
n := UDINT_TO_INT(GVL_Plan.stActive.aSection[nSection].nPointCount);
FOR i := 1 TO n DO
    aCamX[i, 1] := GVL_Plan.stActive.aPoint[nFirst + i - 1].fS_mm;
    aCamX[i, 2] := GVL_Plan.stActive.aPoint[nFirst + i - 1].fU_mm;
    aCamA[i, 1] := GVL_Plan.stActive.aPoint[nFirst + i - 1].fS_mm;
    aCamA[i, 2] := GVL_Plan.stActive.aPoint[nFirst + i - 1].fPhi_deg;
END_FOR
stCamX.pArray := ADR(aCamX);
stCamX.ArraySize := SIZEOF(aCamX);
stCamX.TableType := MC_TableType.MC_TABLETYPE_NONEQUIDISTANT;
stCamX.NoOfRows := INT_TO_UDINT(n);
stCamX.NoOfColumns := 2;
stCamA.pArray := ADR(aCamA);
stCamA.ArraySize := SIZEOF(aCamA);
stCamA.TableType := MC_TableType.MC_TABLETYPE_NONEQUIDISTANT;
stCamA.NoOfRows := INT_TO_UDINT(n);
stCamA.NoOfColumns := 2;
nRotIdx := 1;
bAtRot := FALSE;
bDone := FALSE;
bTableReady := FALSE;
bLoading := TRUE;
bSelExec := FALSE;
fbSelX(Master := GVL_Axis.Z1, Slave := GVL_Axis.X, CamTable := stCamX, Execute := FALSE);
fbSelA(Master := GVL_Axis.Z1, Slave := GVL_Axis.A, CamTable := stCamA, Execute := FALSE);
bSelExec := TRUE;
LoadSection := TRUE;
END_METHOD

METHOD TableReady : BOOL
VAR_INPUT
END_VAR
TableReady := bTableReady AND NOT bLoading;
END_METHOD

METHOD Start : BOOL
VAR_INPUT
END_VAR
IF stStatus.eState = E_KinState.Loaded AND bTableReady THEN
    bInExec := FALSE;
    fbInX(Master := GVL_Axis.Z1, Slave := GVL_Axis.X, Execute := FALSE);
    fbInA(Master := GVL_Axis.Z1, Slave := GVL_Axis.A, Execute := FALSE);
    bHoldPending := FALSE;
    stStatus.eState := E_KinState.Coupling;
    Start := TRUE;
END_IF
END_METHOD

METHOD Hold : BOOL
VAR_INPUT
END_VAR
IF stStatus.eState = E_KinState.Running THEN
    stStatus.eState := E_KinState.Holding;
    Hold := TRUE;
ELSIF stStatus.eState = E_KinState.Coupling THEN
    // noch nicht gefahren: Kopplung fertigstellen lassen, aber nicht losfahren
    bHoldPending := TRUE;
    Hold := TRUE;
END_IF
END_METHOD

METHOD Resume : BOOL
VAR_INPUT
END_VAR
IF stStatus.eState = E_KinState.Held AND NOT bAtRot AND NOT bDone THEN
    stStatus.eState := E_KinState.Running;
    IssueMaster(TRUE);
    Resume := TRUE;
END_IF
END_METHOD

METHOD AtRotation : BOOL
VAR_INPUT
END_VAR
AtRotation := bAtRot AND stStatus.eState = E_KinState.Held;
END_METHOD

METHOD RotationAngle : LREAL
VAR_INPUT
END_VAR
IF nSection >= 1 AND nSection <= GVL_Config.cMaxSections AND nRotIdx >= 1
   AND_THEN nRotIdx <= UINT_TO_INT(GVL_Plan.stActive.aSection[nSection].nRotCount) THEN
    RotationAngle := GVL_Plan.stActive.aSection[nSection].aRot[nRotIdx].fW_deg;
END_IF
END_METHOD

METHOD ContinueAfterRotation : BOOL
VAR_INPUT
END_VAR
IF bAtRot AND stStatus.eState = E_KinState.Held THEN
    bAtRot := FALSE;
    nRotIdx := nRotIdx + 1;
    stStatus.eState := E_KinState.Running;
    IssueMaster(TRUE);
    ContinueAfterRotation := TRUE;
END_IF
END_METHOD

METHOD SectionDone : BOOL
VAR_INPUT
END_VAR
SectionDone := bDone AND stStatus.eState = E_KinState.Held;
END_METHOD

METHOD Abort : BOOL
VAR_INPUT
END_VAR
CASE stStatus.eState OF
E_KinState.Coupling, E_KinState.Running, E_KinState.Holding, E_KinState.Held:
    stStatus.eState := E_KinState.Decoupling;
    nPhase := 0;
    Abort := TRUE;
END_CASE
END_METHOD

METHOD Reset : BOOL
VAR_INPUT
END_VAR
// Nur wenn die Slaves ausgekoppelt sind und keine Achse mehr gestört ist.
IF stStatus.eState = E_KinState.Fault AND nPhase >= 3 THEN
    IF NOT GVL_Devices.aAxis[1].bError AND NOT GVL_Devices.aAxis[3].bError AND NOT GVL_Devices.aAxis[4].bError THEN
        stStatus.bError := FALSE;
        stStatus.nErrorId := 0;
        nPhase := 0;
        bTableReady := FALSE;
        bAtRot := FALSE;
        bDone := FALSE;
        IF GVL_Plan.bValid AND stStatus.nPlanId <> 0 THEN
            stStatus.eState := E_KinState.Loaded;
        ELSE
            stStatus.eState := E_KinState.Idle;
        END_IF
        Reset := TRUE;
    END_IF
END_IF
END_METHOD

METHOD Unload : BOOL
VAR_INPUT
END_VAR
IF stStatus.eState = E_KinState.Idle OR stStatus.eState = E_KinState.Loaded THEN
    stStatus.eState := E_KinState.Idle;
    stStatus.nPlanId := 0;
    nSection := 0;
    bTableReady := FALSE;
    Unload := TRUE;
END_IF
END_METHOD

METHOD IsCoupled : BOOL
VAR_INPUT
END_VAR
CASE stStatus.eState OF
E_KinState.Coupling, E_KinState.Running, E_KinState.Holding, E_KinState.Held, E_KinState.Decoupling:
    IsCoupled := TRUE;
E_KinState.Fault:
    IsCoupled := nPhase < 3;
END_CASE
END_METHOD

METHOD GetStatus : ST_KinStatus
VAR_INPUT
END_VAR
GetStatus := stStatus;
END_METHOD

END_FUNCTION_BLOCK

// ---- 06_HMI/FB_AlarmManager.TcPOU
// Aktive oder nicht quittierte Alarme (max. 32). Texte und Historie liegen im Backend.
// Ein Eintrag verschwindet, wenn die Ursache behoben UND der Alarm quittiert ist.
FUNCTION_BLOCK FB_AlarmManager
VAR_OUTPUT
    nStopCounter : UDINT;     // +1 bei jedem neuen Alarm der Stufe Stop oder Fault (G1 wechselt in Pause)
END_VAR
VAR
    aList : ARRAY[1..32] OF ST_AlarmEntry;
    nCount : INT;
    nChangeCounter : UDINT;
    bOverflow : BOOL;
END_VAR

// Kein zyklischer Anteil; WriteTo() einmal pro Zyklus aufrufen.

METHOD PRIVATE Find : INT
VAR_INPUT
    eCode : E_AlarmCode;
    nSource : DINT;
END_VAR
VAR
    i : INT;
END_VAR
Find := 0;
FOR i := 1 TO nCount DO
    IF aList[i].eCode = eCode AND aList[i].nSource = nSource THEN
        Find := i;
        RETURN;
    END_IF
END_FOR
END_METHOD

METHOD Raise : BOOL
VAR_INPUT
    eCode : E_AlarmCode;
    eSeverity : E_AlarmSeverity;
    nSource : DINT;
    nDetail : UDINT;
END_VAR
VAR
    i : INT;
END_VAR
i := Find(eCode, nSource);
IF i > 0 THEN
    IF aList[i].bActive THEN
        RETURN;           // besteht bereits
    END_IF
ELSE
    IF nCount >= 32 THEN
        bOverflow := TRUE;
        RETURN;
    END_IF
    nCount := nCount + 1;
    i := nCount;
    aList[i].eCode := eCode;
    aList[i].nSource := nSource;
END_IF
aList[i].eSeverity := eSeverity;
aList[i].nDetail := nDetail;
aList[i].nTimestamp := F_GetSystemTime();
aList[i].bActive := TRUE;
aList[i].bAcked := FALSE;
nChangeCounter := nChangeCounter + 1;
IF TO_INT(eSeverity) >= TO_INT(E_AlarmSeverity.Stop) THEN
    nStopCounter := nStopCounter + 1;
END_IF
Raise := TRUE;
END_METHOD

METHOD Clear : BOOL
VAR_INPUT
    eCode : E_AlarmCode;
    nSource : DINT;
    bAnySource : BOOL;
END_VAR
VAR
    i : INT;
END_VAR
FOR i := 1 TO nCount DO
    IF aList[i].eCode = eCode AND (bAnySource OR aList[i].nSource = nSource) AND aList[i].bActive THEN
        aList[i].bActive := FALSE;
        Clear := TRUE;
    END_IF
END_FOR
IF Clear THEN
    nChangeCounter := nChangeCounter + 1;
    Purge();
END_IF
END_METHOD

METHOD Set : BOOL
// Alarm entsprechend einer Bedingung setzen oder zurücknehmen.
VAR_INPUT
    bCondition : BOOL;
    eCode : E_AlarmCode;
    eSeverity : E_AlarmSeverity;
    nSource : DINT;
    nDetail : UDINT;
END_VAR
IF bCondition THEN
    Raise(eCode, eSeverity, nSource, nDetail);
ELSIF IsActive(eCode, nSource, FALSE) THEN
    Clear(eCode, nSource, FALSE);
END_IF
Set := bCondition;
END_METHOD

METHOD Ack : BOOL
VAR_INPUT
    nSlot : DINT;     // 0 = alle
END_VAR
VAR
    i : INT;
END_VAR
FOR i := 1 TO nCount DO
    IF nSlot = 0 OR nSlot = i THEN
        aList[i].bAcked := TRUE;
    END_IF
END_FOR
nChangeCounter := nChangeCounter + 1;
Purge();
Ack := TRUE;
END_METHOD

METHOD PRIVATE Purge
VAR
    i, j : INT;
END_VAR
j := 0;
FOR i := 1 TO nCount DO
    IF aList[i].bActive OR NOT aList[i].bAcked THEN
        j := j + 1;
        IF j <> i THEN
            aList[j] := aList[i];
        END_IF
    END_IF
END_FOR
FOR i := j + 1 TO nCount DO
    aList[i].eCode := E_AlarmCode.None;
    aList[i].eSeverity := E_AlarmSeverity.None;
    aList[i].nSource := 0;
    aList[i].nDetail := 0;
    aList[i].nTimestamp := 0;
    aList[i].bActive := FALSE;
    aList[i].bAcked := FALSE;
END_FOR
nCount := j;
END_METHOD

METHOD IsActive : BOOL
VAR_INPUT
    eCode : E_AlarmCode;
    nSource : DINT;
    bAnySource : BOOL;
END_VAR
VAR
    i : INT;
END_VAR
FOR i := 1 TO nCount DO
    IF aList[i].eCode = eCode AND aList[i].bActive AND (bAnySource OR aList[i].nSource = nSource) THEN
        IsActive := TRUE;
        RETURN;
    END_IF
END_FOR
END_METHOD

METHOD FaultActive : BOOL
// Aktiver Alarm der Stufe Fault.
VAR
    i : INT;
END_VAR
FOR i := 1 TO nCount DO
    IF aList[i].bActive AND aList[i].eSeverity = E_AlarmSeverity.Fault THEN
        FaultActive := TRUE;
        RETURN;
    END_IF
END_FOR
END_METHOD

METHOD WriteTo
VAR_IN_OUT
    stOut : ST_HmiAlarms;
END_VAR
VAR
    i : INT;
    nHigh : INT;
END_VAR
stOut.aEntry := aList;
stOut.nCount := INT_TO_UINT(nCount);
stOut.bOverflow := bOverflow;
stOut.nChangeCounter := nChangeCounter;
nHigh := 0;
stOut.eHighestSeverity := E_AlarmSeverity.None;
FOR i := 1 TO nCount DO
    IF TO_INT(aList[i].eSeverity) > nHigh THEN
        nHigh := TO_INT(aList[i].eSeverity);
        stOut.eHighestSeverity := aList[i].eSeverity;
    END_IF
END_FOR
END_METHOD

END_FUNCTION_BLOCK

